(* Logix 5000 project; controller TFF vendor 1 type 14 code 107 rev 33.11; software revision 33.04; part 7 of 38 *)

        [4,11].DelayTimer.PRE := 2000, [4,11].DelayTimerSP := 2, [4,11].EnableCfg := 1, [4,11].ActiveStateCFg := 1, [4,11].RealInputCfg := 1, [4,11].InputAddressCfg := 11, [4,12].Tag := 'ZS007', [4,12].DelayTimer.PRE := 2000, [4,12].DelayTimerSP := 2, [4,12].EnableCfg := 1, [4,12].ActiveStateCFg := 1, [4,12].RealInputCfg := 1, [4,12].InputAddressCfg := 12, [4,13].Tag := 'ZS008', [4,13].AlarmCurrentValue := 1, [4,13].Override := 1, [4,13].DelayTimer.PRE := 20000, [4,13].DelayTimerSP := 2, [4,13].Priority := 1, [4,13].EnableCfg := 1, [4,13].ActiveStateCFg := 1, [4,13].RealInputCfg := 1, [4,13].InputAddressCfg := 13, [4,13].AlarmCfg := 1, [4,13].OverrideCfg := 1, [4,13].PriorityCfg := 1, [4,13].Cond1Cfg := 1, [4,14].Tag := 'XS011', [4,14].DelayTimer.PRE := 2000, [4,14].DelayTimerSP := 2, [4,14].EnableCfg := 1, [4,14].ActiveStateCFg := 1, [4,14].RealInputCfg := 1, [4,14].InputAddressCfg := 14, [4,15].Tag := 'XS012', [4,15].SoftInput := 1, [4,15].DelayTimer.PRE := 2000, [4,15].DelayTimerSP := 2, [4,15].EnableCfg := 1, [4,15].ActiveStateCFg := 1, [4,15].RealInputCfg := 1, [4,15].InputAddressCfg := 15, [4,16].Tag := 'SIC001DF', [4,16].AlarmCurrentValue := 1, [4,16].Override := 1, [4,16].SoftInput := 1, [4,16].DelayTimer.PRE := 1000, [4,16].DelayTimer.ACC := 3148, [4,16].DelayTimer.EN := 1, [4,16].DelayTimer.DN := 1, [4,16].DelayTimerSP := 1, [4,16].Priority := 1, [4,16].EnableCfg := 1, [4,16].ActiveStateCFg := 1, [4,16].RealInputCfg := 1, [4,16].InputAddressCfg := 16, [4,16].AlarmCfg := 1, [4,16].OverrideCfg := 1, [4,16].PriorityCfg := 1, [4,17].Tag := 'SIC002DF',
        [4,17].AlarmCurrentValue := 1, [4,17].Override := 1, [4,17].SoftInput := 1, [4,17].DelayTimer.PRE := 1000, [4,17].DelayTimer.ACC := 2449345, [4,17].DelayTimer.EN := 1, [4,17].DelayTimer.DN := 1, [4,17].DelayTimerSP := 1, [4,17].Priority := 1, [4,17].EnableCfg := 1, [4,17].ActiveStateCFg := 1, [4,17].RealInputCfg := 1, [4,17].InputAddressCfg := 17, [4,17].AlarmCfg := 1, [4,17].OverrideCfg := 1, [4,17].PriorityCfg := 1, [4,18].Tag := 'AA008', [4,18].AlarmCurrentValue := 1, [4,18].Override := 1, [4,18].DelayTimer.PRE := 1000, [4,18].DelayTimer.ACC := 1042, [4,18].DelayTimer.EN := 1, [4,18].DelayTimer.DN := 1, [4,18].DelayTimerSP := 1, [4,18].Priority := 1, [4,18].EnableCfg := 1, [4,18].ActiveStateCFg := 1, [4,18].RealInputCfg := 1, [4,18].InputAddressCfg := 18, [4,18].AlarmCfg := 1, [4,18].OverrideCfg := 1, [4,18].PriorityCfg := 1, [4,19].Tag := 'LSH001', [4,19].AlarmCurrentValue := 1, [4,19].Override := 1, [4,19].DelayTimer.PRE := 1000, [4,19].DelayTimer.EN := 1, [4,19].DelayTimer.DN := 1, [4,19].DelayTimerSP := 1, [4,19].EnableCfg := 1, [4,19].ActiveStateCFg := 1, [4,19].RealInputCfg := 1, [4,19].InputAddressCfg := 19, [4,19].AlarmCfg := 1, [4,19].OverrideCfg := 1, [4,19].PriorityCfg := 1, [4,20].Tag := 'LSL002', [4,20].AlarmCurrentValue := 1, [4,20].Override := 1, [4,20].DelayTimer.PRE := 1000, [4,20].DelayTimer.EN := 1, [4,20].DelayTimer.DN := 1, [4,20].DelayTimerSP := 1, [4,20].EnableCfg := 1, [4,20].ActiveStateCFg := 1, [4,20].RealInputCfg := 1, [4,20].InputAddressCfg := 20, [4,20].AlarmCfg := 1, [4,20].OverrideCfg := 1, [4,20].PriorityCfg := 1,
        [4,21].Tag := 'PSH001', [4,21].AlarmCurrentValue := 1, [4,21].AlarmAck := 1, [4,21].Alarm := 1, [4,21].Mimic := 5, [4,21].DelayTimer.PRE := 1000, [4,21].DelayTimer.ACC := 1042, [4,21].DelayTimer.EN := 1, [4,21].DelayTimer.DN := 1, [4,21].DelayTimerSP := 1, [4,21].Priority := 1, [4,21].EnableCfg := 1, [4,21].ActiveStateCFg := 1, [4,21].RealInputCfg := 1, [4,21].InputAddressCfg := 21, [4,21].AlarmCfg := 1, [4,21].AlarmONS := 1, [4,22].Tag := 'PSH002', [4,22].AlarmCurrentValue := 1, [4,22].AlarmAck := 1, [4,22].Alarm := 1, [4,22].Mimic := 5, [4,22].DelayTimer.PRE := 1000, [4,22].DelayTimer.ACC := 1042, [4,22].DelayTimer.EN := 1, [4,22].DelayTimer.DN := 1, [4,22].DelayTimerSP := 1, [4,22].Priority := 1, [4,22].EnableCfg := 1, [4,22].ActiveStateCFg := 1, [4,22].RealInputCfg := 1, [4,22].InputAddressCfg := 22, [4,22].AlarmCfg := 1, [4,22].AlarmONS := 1, [4,23].Tag := 'DF48VP001', [4,23].AlarmCurrentValue := 1, [4,23].Override := 1, [4,23].DelayTimer.PRE := 1000, [4,23].DelayTimer.ACC := 1042, [4,23].DelayTimer.EN := 1, [4,23].DelayTimer.DN := 1, [4,23].DelayTimerSP := 1, [4,23].Priority := 1, [4,23].EnableCfg := 1, [4,23].ActiveStateCFg := 1, [4,23].RealInputCfg := 1, [4,23].InputAddressCfg := 23, [4,23].AlarmCfg := 1, [4,23].OverrideCfg := 1, [4,23].PriorityCfg := 1, [4,24].Tag := 'DF48VP002', [4,24].AlarmCurrentValue := 1, [4,24].Override := 1, [4,24].DelayTimer.PRE := 1000, [4,24].DelayTimer.ACC := 1043, [4,24].DelayTimer.EN := 1, [4,24].DelayTimer.DN := 1, [4,24].DelayTimerSP := 1, [4,24].Priority := 1, [4,24].EnableCfg := 1,
        [4,24].ActiveStateCFg := 1, [4,24].RealInputCfg := 1, [4,24].InputAddressCfg := 24, [4,24].AlarmCfg := 1, [4,24].OverrideCfg := 1, [4,24].PriorityCfg := 1, [4,25].Tag := 'XS002', [4,25].AlarmCurrentValue := 1, [4,25].Override := 1, [4,25].DelayTimer.PRE := 20000, [4,25].DelayTimerSP := 2, [4,25].Priority := 1, [4,25].EnableCfg := 1, [4,25].ActiveStateCFg := 1, [4,25].RealInputCfg := 1, [4,25].InputAddressCfg := 25, [4,25].AlarmCfg := 1, [4,25].OverrideCfg := 1, [4,25].PriorityCfg := 1, [4,25].Cond1Cfg := 1, [4,26].Override := 1, [4,26].ActiveStateCFg := 1, [4,26].RealInputCfg := 1, [4,26].InputAddressCfg := 26, [4,26].OverrideCfg := 1, [4,26].PriorityCfg := 1, [4,27].Override := 1, [4,27].SoftInput := 1, [4,27].ActiveStateCFg := 1, [4,27].RealInputCfg := 1, [4,27].InputAddressCfg := 27, [4,27].OverrideCfg := 1, [4,27].PriorityCfg := 1, [4,28].Override := 1, [4,28].SoftInput := 1, [4,28].ActiveStateCFg := 1, [4,28].RealInputCfg := 1, [4,28].InputAddressCfg := 28, [4,28].OverrideCfg := 1, [4,28].PriorityCfg := 1, [4,29].Override := 1, [4,29].SoftInput := 1, [4,29].ActiveStateCFg := 1, [4,29].RealInputCfg := 1, [4,29].InputAddressCfg := 29, [4,29].OverrideCfg := 1, [4,29].PriorityCfg := 1, [4,30].Override := 1, [4,30].SoftInput := 1, [4,30].ActiveStateCFg := 1, [4,30].RealInputCfg := 1, [4,30].InputAddressCfg := 30, [4,30].OverrideCfg := 1, [4,30].PriorityCfg := 1, [4,31].Override := 1, [4,31].ActiveStateCFg := 1, [4,31].RealInputCfg := 1, [4,31].InputAddressCfg := 31, [4,31].OverrideCfg := 1, [4,31].PriorityCfg := 1,
        [4,34].Tag := 'DI1', [4,34].Override := 1, [4,34].SoftInput := 1, [4,34].EnableCfg := 1, [4,34].ActiveStateCFg := 1, [4,34].RealInputCfg := 1, [4,34].InputAddressCfg := 34, [4,34].OverrideCfg := 1, [4,34].PriorityCfg := 1, [4,35].Tag := 'DI2', [4,35].Override := 1, [4,35].EnableCfg := 1, [4,35].ActiveStateCFg := 1, [4,35].RealInputCfg := 1, [4,35].InputAddressCfg := 35, [4,35].OverrideCfg := 1, [4,35].PriorityCfg := 1, [4,36].Tag := 'DI3', [4,36].Override := 1, [4,36].SoftInput := 1, [4,36].EnableCfg := 1, [4,36].ActiveStateCFg := 1, [4,36].RealInputCfg := 1, [4,36].InputAddressCfg := 36, [4,36].OverrideCfg := 1, [4,36].PriorityCfg := 1, [4,37].Tag := 'DI4', [4,37].Override := 1, [4,37].EnableCfg := 1, [4,37].ActiveStateCFg := 1, [4,37].RealInputCfg := 1, [4,37].InputAddressCfg := 37, [4,37].OverrideCfg := 1, [4,37].PriorityCfg := 1, [4,38].Tag := 'DI5', [4,38].Override := 1, [4,38].EnableCfg := 1, [4,38].ActiveStateCFg := 1, [4,38].RealInputCfg := 1, [4,38].InputAddressCfg := 38, [4,38].OverrideCfg := 1, [4,38].PriorityCfg := 1, [4,39].Tag := 'DI6', [4,39].Override := 1, [4,39].SoftInput := 1, [4,39].EnableCfg := 1, [4,39].ActiveStateCFg := 1, [4,39].RealInputCfg := 1, [4,39].InputAddressCfg := 39, [4,39].OverrideCfg := 1, [4,39].PriorityCfg := 1, [4,40].Tag := 'DI7', [4,40].Override := 1, [4,40].EnableCfg := 1, [4,40].ActiveStateCFg := 1, [4,40].RealInputCfg := 1, [4,40].InputAddressCfg := 40, [4,40].OverrideCfg := 1, [4,40].PriorityCfg := 1, [4,41].Tag := 'DI8',
        [4,41].Override := 1, [4,41].EnableCfg := 1, [4,41].ActiveStateCFg := 1, [4,41].RealInputCfg := 1, [4,41].InputAddressCfg := 41, [4,41].OverrideCfg := 1, [4,41].PriorityCfg := 1, [4,50].Tag := 'YA01', [4,50].Desc := 'PC to PLC Com. Failure', [4,50].AlarmCurrentValue := 1, [4,50].Override := 1, [4,50].SoftInput := 1, [4,50].Condition1 := 1, [4,50].Cond1Text := 'HMI HeartBeat received', [4,50].DelayTimer.PRE := 60000, [4,50].DelayTimer.ACC := 598, [4,50].DelayTimer.EN := 1, [4,50].DelayTimer.TT := 1, [4,50].DelayTimerSP := 60, [4,50].EnableCfg := 1, [4,50].InputAddressCfg := 50, [4,50].AlarmCfg := 1, [4,50].AlarmStateCfg := 1, [4,50].OverrideCfg := 1, [4,50].PriorityCfg := 1, [4,50].Cond1Cfg := 1, [4,51].Tag := 'YA02', [4,51].Desc := 'CCP Runtime Com. Failure', [4,51].AlarmCurrentValue := 1, [4,51].Override := 1, [4,51].SoftInput := 1, [4,51].Condition1 := 1, [4,51].Cond1Text := 'HMI HeartBeat received', [4,51].DelayTimer.PRE := 60000, [4,51].DelayTimer.ACC := 60008, [4,51].DelayTimer.EN := 1, [4,51].DelayTimer.DN := 1, [4,51].DelayTimerSP := 60, [4,51].EnableCfg := 1, [4,51].InputAddressCfg := 51, [4,51].AlarmCfg := 1, [4,51].AlarmStateCfg := 1, [4,51].OverrideCfg := 1, [4,51].PriorityCfg := 1, [4,51].Cond1Cfg := 1, [4,52].Tag := 'YA03', [4,52].Desc := 'Hist. Data Collect. Fail', [4,52].AlarmCurrentValue := 1, [4,52].Override := 1, [4,52].SoftInput := 1, [4,52].Condition1 := 1, [4,52].Cond1Text := 'HMI HeartBeat received', [4,52].DelayTimer.PRE := 60000, [4,52].DelayTimer.ACC := 1145, [4,52].DelayTimer.EN := 1, [4,52].DelayTimer.TT := 1, [4,52].DelayTimerSP := 60, [4,52].EnableCfg := 1, [4,52].InputAddressCfg := 52, [4,52].AlarmCfg := 1,
        [4,52].AlarmStateCfg := 1, [4,52].OverrideCfg := 1, [4,52].PriorityCfg := 1, [4,52].Cond1Cfg := 1, [4,53].Tag := 'YA04', [4,53].Desc := 'HDD OverLoad', [4,53].Override := 1, [4,53].DelayTimer.PRE := 60000, [4,53].DelayTimerSP := 60, [4,53].EnableCfg := 1, [4,53].ActiveStateCFg := 1, [4,53].InputAddressCfg := 53, [4,53].AlarmCfg := 1, [4,53].AlarmStateCfg := 1, [4,53].OverrideCfg := 1, [4,53].PriorityCfg := 1, [4,54].Tag := 'YA05', [4,54].Override := 1, [4,54].DelayTimer.PRE := 60000, [4,54].DelayTimerSP := 60, [4,54].EnableCfg := 1, [4,54].ActiveStateCFg := 1, [4,54].InputAddressCfg := 54, [4,54].AlarmCfg := 1, [4,54].AlarmStateCfg := 1, [4,54].OverrideCfg := 1, [4,54].PriorityCfg := 1, [4,55].Tag := 'YA06', [4,55].CurrentValue := 1, [4,55].AlarmCurrentValue := 1, [4,55].Override := 1, [4,55].Mimic := 1, [4,55].SoftInput := 1, [4,55].DelayTimer.PRE := 5000, [4,55].DelayTimer.ACC := 5022, [4,55].DelayTimer.EN := 1, [4,55].DelayTimer.DN := 1, [4,55].DelayTimerSP := 5, [4,55].Priority := 1, [4,55].EnableCfg := 1, [4,55].ActiveStateCFg := 1, [4,55].InputAddressCfg := 55, [4,55].AlarmCfg := 1, [4,55].AlarmStateCfg := 1, [4,55].OverrideCfg := 1, [4,55].PriorityCfg := 1, [4,56].Tag := 'YA07', [4,56].CurrentValue := 1, [4,56].AlarmCurrentValue := 1, [4,56].Override := 1, [4,56].Mimic := 1, [4,56].SoftInput := 1, [4,56].DelayTimer.PRE := 2000, [4,56].DelayTimer.ACC := 2004, [4,56].DelayTimer.EN := 1, [4,56].DelayTimer.DN := 1, [4,56].DelayTimerSP := 2, [4,56].EnableCfg := 1, [4,56].ActiveStateCFg := 1, [4,56].InputAddressCfg := 56,
        [4,56].AlarmCfg := 1, [4,56].AlarmStateCfg := 1, [4,56].OverrideCfg := 1, [4,56].PriorityCfg := 1, [4,57].Tag := 'YA08', [4,57].CurrentValue := 1, [4,57].AlarmCurrentValue := 1, [4,57].Override := 1, [4,57].Mimic := 1, [4,57].SoftInput := 1, [4,57].DelayTimer.PRE := 5000, [4,57].DelayTimer.ACC := 5011, [4,57].DelayTimer.EN := 1, [4,57].DelayTimer.DN := 1, [4,57].DelayTimerSP := 5, [4,57].Priority := 1, [4,57].EnableCfg := 1, [4,57].ActiveStateCFg := 1, [4,57].InputAddressCfg := 57, [4,57].AlarmCfg := 1, [4,57].AlarmStateCfg := 1, [4,57].OverrideCfg := 1, [4,57].PriorityCfg := 1, [4,58].Tag := 'YA09', [4,58].CurrentValue := 1, [4,58].AlarmCurrentValue := 1, [4,58].Override := 1, [4,58].Mimic := 1, [4,58].SoftInput := 1, [4,58].DelayTimer.PRE := 2000, [4,58].DelayTimer.ACC := 2050, [4,58].DelayTimer.EN := 1, [4,58].DelayTimer.DN := 1, [4,58].DelayTimerSP := 2, [4,58].EnableCfg := 1, [4,58].ActiveStateCFg := 1, [4,58].InputAddressCfg := 58, [4,58].AlarmCfg := 1, [4,58].AlarmStateCfg := 1, [4,58].OverrideCfg := 1, [4,58].PriorityCfg := 1, [4,59].Tag := 'YA10', [4,59].CurrentValue := 1, [4,59].Mimic := 1, [4,59].Priority := 1, [4,59].EnableCfg := 1, [4,59].InputAddressCfg := 59, [4,59].AlarmCfg := 1, [4,59].AlarmStateCfg := 1, [4,60].Tag := 'YA11', [4,60].AlarmCurrentValue := 1, [4,60].Override := 1, [4,60].DelayTimer.PRE := 5000, [4,60].DelayTimer.ACC := 5010, [4,60].DelayTimer.EN := 1, [4,60].DelayTimer.DN := 1, [4,60].DelayTimerSP := 5, [4,60].EnableCfg := 1, [4,60].ActiveStateCFg := 1, [4,60].InputAddressCfg := 60,
        [4,60].AlarmCfg := 1, [4,60].OverrideCfg := 1, [4,60].PriorityCfg := 1, [4,61].Tag := 'YA12', [4,61].Override := 1, [4,61].DelayTimer.PRE := 2000, [4,61].DelayTimerSP := 2, [4,61].EnableCfg := 1, [4,61].ActiveStateCFg := 1, [4,61].InputAddressCfg := 61, [4,61].AlarmCfg := 1, [4,61].AlarmStateCfg := 1, [4,61].OverrideCfg := 1, [4,61].PriorityCfg := 1, [4,62].Tag := 'UserNCr1', [4,62].CurrentValue := 1, [4,62].Mimic := 1, [4,62].EnableCfg := 1, [4,62].InputAddressCfg := 62, [4,63].Tag := 'UserCr1', [4,63].SoftInput := 1, [4,63].Priority := 1, [4,63].EnableCfg := 1, [4,63].InputAddressCfg := 63, [4,64].Tag := 'UserNCr2', [4,64].CurrentValue := 1, [4,64].Mimic := 1, [4,64].EnableCfg := 1, [4,64].InputAddressCfg := 64, [4,65].Tag := 'UserCr2', [4,65].CurrentValue := 1, [4,65].Mimic := 1, [4,65].Priority := 1, [4,65].EnableCfg := 1, [4,65].InputAddressCfg := 65, [4,66].Tag := 'LV001_Err', [4,66].Override := 1, [4,66].DelayTimer.PRE := 2000, [4,66].DelayTimerSP := 2, [4,66].EnableCfg := 1, [4,66].ActiveStateCFg := 1, [4,66].InputAddressCfg := 66, [4,66].AlarmCfg := 1, [4,66].AlarmStateCfg := 1, [4,66].OverrideCfg := 1, [4,66].PriorityCfg := 1, [4,67].Tag := 'LV002_Err', [4,67].Override := 1, [4,67].DelayTimer.PRE := 2000, [4,67].DelayTimerSP := 2, [4,67].EnableCfg := 1, [4,67].ActiveStateCFg := 1, [4,67].InputAddressCfg := 67, [4,67].AlarmCfg := 1, [4,67].AlarmStateCfg := 1, [4,67].OverrideCfg := 1, [4,67].PriorityCfg := 1, [4,68].CurrentValue := 1, [4,68].AlarmCurrentValue := 1, [4,68].Override := 1,
        [4,68].Mimic := 1, [4,68].SoftInput := 1, [4,68].DelayTimer.PRE := 1000, [4,68].DelayTimer.ACC := 3526, [4,68].DelayTimer.EN := 1, [4,68].DelayTimer.DN := 1, [4,68].DelayTimerSP := 1, [4,68].Priority := 1, [4,68].EnableCfg := 1, [4,68].ActiveStateCFg := 1, [4,68].InputAddressCfg := 68, [4,68].AlarmCfg := 1, [4,68].AlarmStateCfg := 1, [4,68].OverrideCfg := 1, [4,69].Override := 1, [4,69].EnableCfg := 1, [4,69].ActiveStateCFg := 1, [4,69].InputAddressCfg := 69, [4,69].AlarmCfg := 1, [4,69].AlarmStateCfg := 1, [4,69].OverrideCfg := 1, [4,69].PriorityCfg := 1, [4,70].CurrentValue := 1, [4,70].Mimic := 1, [4,70].DelayTimer.PRE := 2000, [4,70].DelayTimerSP := 2, [4,70].Priority := 1, [4,70].ActiveStateCFg := 1, [4,70].InputAddressCfg := 70, [4,70].AlarmStateCfg := 1, [4,70].OverrideCfg := 1, [4,70].PriorityCfg := 1, [4,71].CurrentValue := 1, [4,71].AlarmCurrentValue := 1, [4,71].AlarmAck := 1, [4,71].Mimic := 5, [4,71].DelayTimer.PRE := 2000, [4,71].DelayTimer.ACC := 2053, [4,71].DelayTimer.EN := 1, [4,71].DelayTimer.DN := 1, [4,71].DelayTimerSP := 2, [4,71].Priority := 1, [4,71].ActiveStateCFg := 1, [4,71].InputAddressCfg := 71, [4,71].AlarmStateCfg := 1, [4,71].OverrideCfg := 1, [4,71].PriorityCfg := 1, [4,71].AlarmONS := 1, [4,72].CurrentValue := 1, [4,72].Mimic := 1, [4,72].DelayTimer.PRE := 2000, [4,72].DelayTimerSP := 2, [4,72].ActiveStateCFg := 1, [4,72].InputAddressCfg := 72, [4,72].AlarmStateCfg := 1, [4,72].OverrideCfg := 1, [4,72].PriorityCfg := 1, [4,73].CurrentValue := 1, [4,73].Mimic := 1, [4,73].DelayTimer.PRE := 2000,
        [4,73].DelayTimerSP := 2, [4,73].ActiveStateCFg := 1, [4,73].InputAddressCfg := 73, [4,73].AlarmStateCfg := 1, [4,73].OverrideCfg := 1, [4,73].PriorityCfg := 1, [4,74].CurrentValue := 1, [4,74].Mimic := 1, [4,74].DelayTimer.PRE := 2000, [4,74].DelayTimerSP := 2, [4,74].ActiveStateCFg := 1, [4,74].InputAddressCfg := 74, [4,74].AlarmStateCfg := 1, [4,74].OverrideCfg := 1, [4,74].PriorityCfg := 1, [4,75].CurrentValue := 1, [4,75].AlarmCurrentValue := 1, [4,75].AlarmAck := 1, [4,75].Alarm := 1, [4,75].Mimic := 3, [4,75].SoftInput := 1, [4,75].DelayTimer.PRE := 2000, [4,75].DelayTimer.ACC := 44, [4,75].DelayTimer.EN := 1, [4,75].DelayTimer.DN := 1, [4,75].DelayTimerSP := 2, [4,75].ActiveStateCFg := 1, [4,75].InputAddressCfg := 75, [4,75].AlarmStateCfg := 1, [4,75].OverrideCfg := 1, [4,75].PriorityCfg := 1, [4,75].AlarmONS := 1, [4,76].CurrentValue := 1, [4,76].Mimic := 1, [4,76].DelayTimer.PRE := 2000, [4,76].DelayTimerSP := 2, [4,76].Priority := 1, [4,76].ActiveStateCFg := 1, [4,76].InputAddressCfg := 76, [4,76].AlarmStateCfg := 1, [4,76].OverrideCfg := 1, [4,76].PriorityCfg := 1, [4,77].CurrentValue := 1, [4,77].Mimic := 1, [4,77].DelayTimer.PRE := 2000, [4,77].DelayTimerSP := 2, [4,77].Priority := 1, [4,77].ActiveStateCFg := 1, [4,77].InputAddressCfg := 77, [4,77].AlarmStateCfg := 1, [4,77].OverrideCfg := 1, [4,77].PriorityCfg := 1, [4,78].CurrentValue := 1, [4,78].AlarmCurrentValue := 1, [4,78].AlarmAck := 1, [4,78].Alarm := 1, [4,78].Mimic := 5, [4,78].SoftInput := 1, [4,78].DelayTimer.PRE := 2000, [4,78].DelayTimer.ACC := 45,
        [4,78].DelayTimer.EN := 1, [4,78].DelayTimer.DN := 1, [4,78].DelayTimerSP := 2, [4,78].Priority := 1, [4,78].ActiveStateCFg := 1, [4,78].InputAddressCfg := 78, [4,78].AlarmStateCfg := 1, [4,78].OverrideCfg := 1, [4,78].PriorityCfg := 1, [4,78].AlarmONS := 1, [4,79].CurrentValue := 1, [4,79].AlarmCurrentValue := 1, [4,79].Mimic := 1, [4,79].DelayTimer.PRE := 2000, [4,79].DelayTimer.ACC := 44, [4,79].DelayTimer.EN := 1, [4,79].DelayTimer.DN := 1, [4,79].DelayTimerSP := 2, [4,79].Priority := 1, [4,79].ActiveStateCFg := 1, [4,79].InputAddressCfg := 79, [4,79].AlarmStateCfg := 1, [4,79].OverrideCfg := 1, [4,79].PriorityCfg := 1, [4,80].CurrentValue := 1, [4,80].AlarmCurrentValue := 1, [4,80].Mimic := 1, [4,80].DelayTimer.PRE := 2000, [4,80].DelayTimer.ACC := 44, [4,80].DelayTimer.EN := 1, [4,80].DelayTimer.DN := 1, [4,80].DelayTimerSP := 2, [4,80].Priority := 1, [4,80].ActiveStateCFg := 1, [4,80].InputAddressCfg := 80, [4,80].AlarmStateCfg := 1, [4,80].OverrideCfg := 1, [4,80].PriorityCfg := 1, [4,81].CurrentValue := 1, [4,81].AlarmCurrentValue := 1, [4,81].Mimic := 1, [4,81].DelayTimer.PRE := 2000, [4,81].DelayTimer.ACC := 44, [4,81].DelayTimer.EN := 1, [4,81].DelayTimer.DN := 1, [4,81].DelayTimerSP := 2, [4,81].ActiveStateCFg := 1, [4,81].InputAddressCfg := 81, [4,81].AlarmStateCfg := 1, [4,81].OverrideCfg := 1, [4,81].PriorityCfg := 1, [4,82].CurrentValue := 1, [4,82].AlarmCurrentValue := 1, [4,82].Mimic := 1, [4,82].DelayTimer.PRE := 2000, [4,82].DelayTimer.ACC := 44, [4,82].DelayTimer.EN := 1, [4,82].DelayTimer.DN := 1, [4,82].DelayTimerSP := 2, [4,82].Priority := 1,
        [4,82].ActiveStateCFg := 1, [4,82].InputAddressCfg := 82, [4,82].AlarmStateCfg := 1, [4,82].OverrideCfg := 1, [4,82].PriorityCfg := 1, [4,83].CurrentValue := 1, [4,83].AlarmCurrentValue := 1, [4,83].AlarmAck := 1, [4,83].Alarm := 1, [4,83].Mimic := 5, [4,83].SoftInput := 1, [4,83].DelayTimer.PRE := 2000, [4,83].DelayTimer.ACC := 44, [4,83].DelayTimer.EN := 1, [4,83].DelayTimer.DN := 1, [4,83].DelayTimerSP := 2, [4,83].Priority := 1, [4,83].ActiveStateCFg := 1, [4,83].InputAddressCfg := 83, [4,83].AlarmStateCfg := 1, [4,83].OverrideCfg := 1, [4,83].PriorityCfg := 1, [4,83].AlarmONS := 1, [4,84].CurrentValue := 1, [4,84].Mimic := 1, [4,84].DelayTimer.PRE := 2000, [4,84].DelayTimerSP := 2, [4,84].Priority := 1, [4,84].ActiveStateCFg := 1, [4,84].InputAddressCfg := 84, [4,84].AlarmStateCfg := 1, [4,84].OverrideCfg := 1, [4,84].PriorityCfg := 1, [4,85].CurrentValue := 1, [4,85].AlarmCurrentValue := 1, [4,85].AlarmAck := 1, [4,85].Alarm := 1, [4,85].Mimic := 3, [4,85].SoftInput := 1, [4,85].DelayTimer.PRE := 2000, [4,85].DelayTimer.ACC := 2021, [4,85].DelayTimer.EN := 1, [4,85].DelayTimer.DN := 1, [4,85].DelayTimerSP := 2, [4,85].ActiveStateCFg := 1, [4,85].InputAddressCfg := 85, [4,85].AlarmStateCfg := 1, [4,85].OverrideCfg := 1, [4,85].PriorityCfg := 1, [4,85].AlarmONS := 1, [4,86].CurrentValue := 1, [4,86].Mimic := 1, [4,86].DelayTimer.PRE := 2000, [4,86].DelayTimerSP := 2, [4,86].ActiveStateCFg := 1, [4,86].InputAddressCfg := 86, [4,86].AlarmStateCfg := 1, [4,86].OverrideCfg := 1, [4,86].PriorityCfg := 1, [4,87].CurrentValue := 1,
        [4,87].Mimic := 1, [4,87].DelayTimer.PRE := 2000, [4,87].DelayTimerSP := 2, [4,87].ActiveStateCFg := 1, [4,87].InputAddressCfg := 87, [4,87].AlarmStateCfg := 1, [4,87].OverrideCfg := 1, [4,87].PriorityCfg := 1, [4,88].CurrentValue := 1, [4,88].Mimic := 1, [4,88].DelayTimer.PRE := 2000, [4,88].DelayTimerSP := 2, [4,88].ActiveStateCFg := 1, [4,88].InputAddressCfg := 88, [4,88].AlarmStateCfg := 1, [4,88].OverrideCfg := 1, [4,88].PriorityCfg := 1, [4,89].CurrentValue := 1, [4,89].Mimic := 1, [4,89].DelayTimer.PRE := 2000, [4,89].DelayTimerSP := 2, [4,89].ActiveStateCFg := 1, [4,89].InputAddressCfg := 89, [4,89].AlarmStateCfg := 1, [4,89].OverrideCfg := 1, [4,89].PriorityCfg := 1, [4,90].Tag := 'PI001_SIG', [4,90].CurrentValue := 1, [4,90].AlarmCurrentValue := 1, [4,90].AlarmAck := 1, [4,90].Alarm := 1, [4,90].Mimic := 5, [4,90].SoftInput := 1, [4,90].DelayTimer.PRE := 2000, [4,90].DelayTimer.ACC := 6308, [4,90].DelayTimer.EN := 1, [4,90].DelayTimer.DN := 1, [4,90].DelayTimerSP := 2, [4,90].Priority := 1, [4,90].EnableCfg := 1, [4,90].ActiveStateCFg := 1, [4,90].InputAddressCfg := 90, [4,90].AlarmCfg := 1, [4,90].AlarmStateCfg := 1, [4,90].OverrideCfg := 1, [4,90].PriorityCfg := 1, [4,90].AlarmONS := 1, [4,91].Tag := 'FI001_SIG', [4,91].CurrentValue := 1, [4,91].AlarmCurrentValue := 1, [4,91].AlarmAck := 1, [4,91].Alarm := 1, [4,91].Mimic := 5, [4,91].SoftInput := 1, [4,91].DelayTimer.PRE := 2000, [4,91].DelayTimer.ACC := 2025, [4,91].DelayTimer.EN := 1, [4,91].DelayTimer.DN := 1, [4,91].DelayTimerSP := 2, [4,91].Priority := 1,
        [4,91].EnableCfg := 1, [4,91].ActiveStateCFg := 1, [4,91].InputAddressCfg := 91, [4,91].AlarmCfg := 1, [4,91].AlarmStateCfg := 1, [4,91].OverrideCfg := 1, [4,91].PriorityCfg := 1, [4,91].AlarmONS := 1, [4,92].Tag := 'PI002_SIG', [4,92].CurrentValue := 1, [4,92].AlarmCurrentValue := 1, [4,92].AlarmAck := 1, [4,92].Alarm := 1, [4,92].Mimic := 5, [4,92].SoftInput := 1, [4,92].DelayTimer.PRE := 2000, [4,92].DelayTimer.EN := 1, [4,92].DelayTimer.DN := 1, [4,92].DelayTimerSP := 2, [4,92].Priority := 1, [4,92].EnableCfg := 1, [4,92].ActiveStateCFg := 1, [4,92].InputAddressCfg := 92, [4,92].AlarmCfg := 1, [4,92].AlarmStateCfg := 1, [4,92].OverrideCfg := 1, [4,92].PriorityCfg := 1, [4,92].AlarmONS := 1, [4,93].Tag := 'FI002_SIG', [4,93].CurrentValue := 1, [4,93].AlarmCurrentValue := 1, [4,93].AlarmAck := 1, [4,93].Alarm := 1, [4,93].Mimic := 5, [4,93].SoftInput := 1, [4,93].DelayTimer.PRE := 2000, [4,93].DelayTimer.ACC := 2049, [4,93].DelayTimer.EN := 1, [4,93].DelayTimer.DN := 1, [4,93].DelayTimerSP := 2, [4,93].Priority := 1, [4,93].EnableCfg := 1, [4,93].ActiveStateCFg := 1, [4,93].InputAddressCfg := 93, [4,93].AlarmCfg := 1, [4,93].AlarmStateCfg := 1, [4,93].OverrideCfg := 1, [4,93].PriorityCfg := 1, [4,93].AlarmONS := 1, [4,94].Tag := 'PI003_SIG', [4,94].CurrentValue := 1, [4,94].AlarmCurrentValue := 1, [4,94].AlarmAck := 1, [4,94].Alarm := 1, [4,94].Mimic := 3, [4,94].SoftInput := 1, [4,94].DelayTimer.PRE := 2000, [4,94].DelayTimer.ACC := 37, [4,94].DelayTimer.EN := 1, [4,94].DelayTimer.DN := 1,
        [4,94].DelayTimerSP := 2, [4,94].EnableCfg := 1, [4,94].ActiveStateCFg := 1, [4,94].InputAddressCfg := 94, [4,94].AlarmCfg := 1, [4,94].AlarmStateCfg := 1, [4,94].OverrideCfg := 1, [4,94].PriorityCfg := 1, [4,94].AlarmONS := 1, [4,95].Tag := 'AI102_SIG', [4,95].CurrentValue := 1, [4,95].AlarmCurrentValue := 1, [4,95].AlarmAck := 1, [4,95].Alarm := 1, [4,95].Mimic := 5, [4,95].SoftInput := 1, [4,95].DelayTimer.PRE := 2000, [4,95].DelayTimer.ACC := 3550, [4,95].DelayTimer.EN := 1, [4,95].DelayTimer.DN := 1, [4,95].DelayTimerSP := 2, [4,95].Priority := 1, [4,95].EnableCfg := 1, [4,95].ActiveStateCFg := 1, [4,95].InputAddressCfg := 95, [4,95].AlarmCfg := 1, [4,95].AlarmStateCfg := 1, [4,95].OverrideCfg := 1, [4,95].PriorityCfg := 1, [4,95].AlarmONS := 1, [4,96].Tag := 'AI103_SIG', [4,96].CurrentValue := 1, [4,96].AlarmCurrentValue := 1, [4,96].AlarmAck := 1, [4,96].Alarm := 1, [4,96].Mimic := 5, [4,96].SoftInput := 1, [4,96].DelayTimer.PRE := 2000, [4,96].DelayTimer.EN := 1, [4,96].DelayTimer.DN := 1, [4,96].DelayTimerSP := 2, [4,96].Priority := 1, [4,96].EnableCfg := 1, [4,96].ActiveStateCFg := 1, [4,96].InputAddressCfg := 96, [4,96].AlarmCfg := 1, [4,96].AlarmStateCfg := 1, [4,96].OverrideCfg := 1, [4,96].PriorityCfg := 1, [4,96].AlarmONS := 1, [4,97].Tag := 'AI201A_SIG', [4,97].CurrentValue := 1, [4,97].AlarmCurrentValue := 1, [4,97].AlarmAck := 1, [4,97].Alarm := 1, [4,97].Mimic := 5, [4,97].SoftInput := 1, [4,97].DelayTimer.PRE := 2000, [4,97].DelayTimer.EN := 1, [4,97].DelayTimer.DN := 1,
        [4,97].DelayTimerSP := 2, [4,97].Priority := 1, [4,97].EnableCfg := 1, [4,97].ActiveStateCFg := 1, [4,97].InputAddressCfg := 97, [4,97].AlarmCfg := 1, [4,97].AlarmStateCfg := 1, [4,97].OverrideCfg := 1, [4,97].PriorityCfg := 1, [4,97].AlarmONS := 1, [4,98].Tag := 'AI201B_SIG', [4,98].CurrentValue := 1, [4,98].AlarmCurrentValue := 1, [4,98].AlarmAck := 1, [4,98].Alarm := 1, [4,98].Mimic := 5, [4,98].SoftInput := 1, [4,98].DelayTimer.PRE := 2000, [4,98].DelayTimer.EN := 1, [4,98].DelayTimer.DN := 1, [4,98].DelayTimerSP := 2, [4,98].Priority := 1, [4,98].EnableCfg := 1, [4,98].ActiveStateCFg := 1, [4,98].InputAddressCfg := 98, [4,98].AlarmCfg := 1, [4,98].AlarmStateCfg := 1, [4,98].OverrideCfg := 1, [4,98].PriorityCfg := 1, [4,98].AlarmONS := 1, [4,99].Tag := 'TI201_SIG', [4,99].CurrentValue := 1, [4,99].AlarmCurrentValue := 1, [4,99].AlarmAck := 1, [4,99].Alarm := 1, [4,99].Mimic := 3, [4,99].SoftInput := 1, [4,99].DelayTimer.PRE := 2000, [4,99].DelayTimer.EN := 1, [4,99].DelayTimer.DN := 1, [4,99].DelayTimerSP := 2, [4,99].EnableCfg := 1, [4,99].ActiveStateCFg := 1, [4,99].InputAddressCfg := 99, [4,99].AlarmCfg := 1, [4,99].AlarmStateCfg := 1, [4,99].OverrideCfg := 1, [4,99].PriorityCfg := 1, [4,99].AlarmONS := 1, [4,100].Tag := 'AI202_SIG', [4,100].CurrentValue := 1, [4,100].AlarmCurrentValue := 1, [4,100].AlarmAck := 1, [4,100].Alarm := 1, [4,100].Mimic := 5, [4,100].SoftInput := 1, [4,100].DelayTimer.PRE := 2000, [4,100].DelayTimer.EN := 1, [4,100].DelayTimer.DN := 1, [4,100].DelayTimerSP := 2,
        [4,100].Priority := 1, [4,100].EnableCfg := 1, [4,100].ActiveStateCFg := 1, [4,100].InputAddressCfg := 100, [4,100].AlarmCfg := 1, [4,100].AlarmStateCfg := 1, [4,100].OverrideCfg := 1, [4,100].PriorityCfg := 1, [4,100].AlarmONS := 1, [4,101].Tag := 'AI203_SIG', [4,101].CurrentValue := 1, [4,101].AlarmCurrentValue := 1, [4,101].AlarmAck := 1, [4,101].Alarm := 1, [4,101].Mimic := 5, [4,101].SoftInput := 1, [4,101].DelayTimer.PRE := 2000, [4,101].DelayTimer.EN := 1, [4,101].DelayTimer.DN := 1, [4,101].DelayTimerSP := 2, [4,101].Priority := 1, [4,101].EnableCfg := 1, [4,101].ActiveStateCFg := 1, [4,101].InputAddressCfg := 101, [4,101].AlarmCfg := 1, [4,101].AlarmStateCfg := 1, [4,101].OverrideCfg := 1, [4,101].PriorityCfg := 1, [4,101].AlarmONS := 1, [4,102].Tag := 'AI204_SIG', [4,102].CurrentValue := 1, [4,102].AlarmCurrentValue := 1, [4,102].AlarmAck := 1, [4,102].Alarm := 1, [4,102].Mimic := 5, [4,102].SoftInput := 1, [4,102].DelayTimer.PRE := 2000, [4,102].DelayTimer.EN := 1, [4,102].DelayTimer.DN := 1, [4,102].DelayTimerSP := 2, [4,102].Priority := 1, [4,102].EnableCfg := 1, [4,102].ActiveStateCFg := 1, [4,102].InputAddressCfg := 102, [4,102].AlarmCfg := 1, [4,102].AlarmStateCfg := 1, [4,102].OverrideCfg := 1, [4,102].PriorityCfg := 1, [4,102].AlarmONS := 1, [4,103].Tag := 'PCV032_SIG', [4,103].CurrentValue := 1, [4,103].AlarmCurrentValue := 1, [4,103].AlarmAck := 1, [4,103].Alarm := 1, [4,103].Mimic := 5, [4,103].SoftInput := 1, [4,103].DelayTimer.PRE := 2000, [4,103].DelayTimer.ACC := 4119948, [4,103].DelayTimer.EN := 1, [4,103].DelayTimer.DN := 1,
        [4,103].DelayTimerSP := 2, [4,103].Priority := 1, [4,103].EnableCfg := 1, [4,103].ActiveStateCFg := 1, [4,103].InputAddressCfg := 103, [4,103].AlarmCfg := 1, [4,103].AlarmStateCfg := 1, [4,103].OverrideCfg := 1, [4,103].PriorityCfg := 1, [4,103].AlarmONS := 1, [5,0].Tag := 'PISL601', [5,0].AlarmCurrentValue := 1, [5,0].Override := 1, [5,0].DelayTimer.PRE := 2000, [5,0].DelayTimer.ACC := 129444, [5,0].DelayTimer.EN := 1, [5,0].DelayTimer.DN := 1, [5,0].DelayTimerSP := 2, [5,0].Priority := 1, [5,0].EnableCfg := 1, [5,0].ActiveStateCFg := 1, [5,0].RealInputCfg := 1, [5,0].AlarmCfg := 1, [5,0].OverrideCfg := 1, [5,0].PriorityCfg := 1, [5,1].Tag := 'PISL602', [5,1].AlarmCurrentValue := 1, [5,1].Override := 1, [5,1].Condition2 := 1, [5,1].DelayTimer.PRE := 2000, [5,1].DelayTimer.ACC := 44686, [5,1].DelayTimer.EN := 1, [5,1].DelayTimer.DN := 1, [5,1].DelayTimerSP := 2, [5,1].Priority := 1, [5,1].EnableCfg := 1, [5,1].ActiveStateCFg := 1, [5,1].RealInputCfg := 1, [5,1].InputAddressCfg := 1, [5,1].AlarmCfg := 1, [5,1].OverrideCfg := 1, [5,1].PriorityCfg := 1, [5,2].Tag := 'ES001', [5,2].CurrentValue := 1, [5,2].Mimic := 1, [5,2].DelayTimer.PRE := 1000, [5,2].DelayTimerSP := 1, [5,2].Priority := 1, [5,2].EnableCfg := 1, [5,2].ActiveStateCFg := 1, [5,2].RealInputCfg := 1, [5,2].InputAddressCfg := 2, [5,2].AlarmCfg := 1, [5,3].Tag := 'RSBUZZ', [5,3].DelayTimer.PRE := 2000, [5,3].DelayTimerSP := 2, [5,3].EnableCfg := 1, [5,3].ActiveStateCFg := 1, [5,3].RealInputCfg := 1, [5,3].InputAddressCfg := 3,
        [5,4].Tag := 'DF24VDC', [5,4].AlarmCurrentValue := 1, [5,4].Override := 1, [5,4].DelayTimer.PRE := 1000, [5,4].DelayTimer.ACC := 11063, [5,4].DelayTimer.EN := 1, [5,4].DelayTimer.DN := 1, [5,4].DelayTimerSP := 1, [5,4].Priority := 1, [5,4].EnableCfg := 1, [5,4].ActiveStateCFg := 1, [5,4].RealInputCfg := 1, [5,4].InputAddressCfg := 4, [5,4].AlarmCfg := 1, [5,4].OverrideCfg := 1, [5,4].PriorityCfg := 1, [5,5].Tag := 'ZS008', [5,5].AlarmCurrentValue := 1, [5,5].Override := 1, [5,5].DelayTimer.PRE := 1000, [5,5].DelayTimer.ACC := 1072, [5,5].DelayTimer.EN := 1, [5,5].DelayTimer.DN := 1, [5,5].DelayTimerSP := 1, [5,5].Priority := 1, [5,5].EnableCfg := 1, [5,5].ActiveStateCFg := 1, [5,5].RealInputCfg := 1, [5,5].InputAddressCfg := 5, [5,5].AlarmCfg := 1, [5,5].OverrideCfg := 1, [5,6].Tag := 'ZS001', [5,6].DelayTimer.PRE := 2000, [5,6].DelayTimerSP := 2, [5,6].EnableCfg := 1, [5,6].ActiveStateCFg := 1, [5,6].RealInputCfg := 1, [5,6].InputAddressCfg := 6, [5,7].Tag := 'ZS002', [5,7].DelayTimer.PRE := 2000, [5,7].DelayTimerSP := 2, [5,7].EnableCfg := 1, [5,7].ActiveStateCFg := 1, [5,7].RealInputCfg := 1, [5,7].InputAddressCfg := 7, [5,8].Tag := 'ZS003', [5,8].DelayTimer.PRE := 2000, [5,8].DelayTimerSP := 2, [5,8].EnableCfg := 1, [5,8].ActiveStateCFg := 1, [5,8].RealInputCfg := 1, [5,8].InputAddressCfg := 8, [5,9].Tag := 'ZS004', [5,9].DelayTimer.PRE := 2000, [5,9].DelayTimerSP := 2, [5,9].EnableCfg := 1, [5,9].ActiveStateCFg := 1, [5,9].RealInputCfg := 1, [5,9].InputAddressCfg := 9, [5,10].Tag := 'ZS005',
        [5,10].DelayTimer.PRE := 2000, [5,10].DelayTimerSP := 2, [5,10].EnableCfg := 1, [5,10].ActiveStateCFg := 1, [5,10].RealInputCfg := 1, [5,10].InputAddressCfg := 10, [5,11].Tag := 'ZS006', [5,11].DelayTimer.PRE := 2000, [5,11].DelayTimerSP := 2, [5,11].EnableCfg := 1, [5,11].ActiveStateCFg := 1, [5,11].RealInputCfg := 1, [5,11].InputAddressCfg := 11, [5,12].Tag := 'ZS007', [5,12].DelayTimer.PRE := 2000, [5,12].DelayTimerSP := 2, [5,12].EnableCfg := 1, [5,12].ActiveStateCFg := 1, [5,12].RealInputCfg := 1, [5,12].InputAddressCfg := 12, [5,13].Tag := 'ZS008', [5,13].AlarmCurrentValue := 1, [5,13].Override := 1, [5,13].DelayTimer.PRE := 20000, [5,13].DelayTimerSP := 2, [5,13].Priority := 1, [5,13].EnableCfg := 1, [5,13].ActiveStateCFg := 1, [5,13].RealInputCfg := 1, [5,13].InputAddressCfg := 13, [5,13].AlarmCfg := 1, [5,13].OverrideCfg := 1, [5,13].PriorityCfg := 1, [5,13].Cond1Cfg := 1, [5,14].Tag := 'XS011', [5,14].DelayTimer.PRE := 2000, [5,14].DelayTimerSP := 2, [5,14].EnableCfg := 1, [5,14].ActiveStateCFg := 1, [5,14].RealInputCfg := 1, [5,14].InputAddressCfg := 14, [5,15].Tag := 'XS012', [5,15].SoftInput := 1, [5,15].DelayTimer.PRE := 2000, [5,15].DelayTimerSP := 2, [5,15].EnableCfg := 1, [5,15].ActiveStateCFg := 1, [5,15].RealInputCfg := 1, [5,15].InputAddressCfg := 15, [5,16].Tag := 'SIC001DF', [5,16].AlarmCurrentValue := 1, [5,16].Override := 1, [5,16].SoftInput := 1, [5,16].DelayTimer.PRE := 1000, [5,16].DelayTimer.ACC := 3148, [5,16].DelayTimer.EN := 1, [5,16].DelayTimer.DN := 1, [5,16].DelayTimerSP := 1, [5,16].Priority := 1, [5,16].EnableCfg := 1,
        [5,16].ActiveStateCFg := 1, [5,16].RealInputCfg := 1, [5,16].InputAddressCfg := 16, [5,16].AlarmCfg := 1, [5,16].OverrideCfg := 1, [5,16].PriorityCfg := 1, [5,17].Tag := 'SIC002DF', [5,17].AlarmCurrentValue := 1, [5,17].Override := 1, [5,17].SoftInput := 1, [5,17].DelayTimer.PRE := 1000, [5,17].DelayTimer.ACC := 2449345, [5,17].DelayTimer.EN := 1, [5,17].DelayTimer.DN := 1, [5,17].DelayTimerSP := 1, [5,17].Priority := 1, [5,17].EnableCfg := 1, [5,17].ActiveStateCFg := 1, [5,17].RealInputCfg := 1, [5,17].InputAddressCfg := 17, [5,17].AlarmCfg := 1, [5,17].OverrideCfg := 1, [5,17].PriorityCfg := 1, [5,18].Tag := 'AA008', [5,18].AlarmCurrentValue := 1, [5,18].Override := 1, [5,18].DelayTimer.PRE := 1000, [5,18].DelayTimer.EN := 1, [5,18].DelayTimer.DN := 1, [5,18].DelayTimerSP := 1, [5,18].Priority := 1, [5,18].EnableCfg := 1, [5,18].ActiveStateCFg := 1, [5,18].RealInputCfg := 1, [5,18].InputAddressCfg := 18, [5,18].AlarmCfg := 1, [5,18].OverrideCfg := 1, [5,18].PriorityCfg := 1, [5,19].Tag := 'LSH001', [5,19].AlarmCurrentValue := 1, [5,19].Override := 1, [5,19].DelayTimer.PRE := 1000, [5,19].DelayTimer.EN := 1, [5,19].DelayTimer.DN := 1, [5,19].DelayTimerSP := 1, [5,19].EnableCfg := 1, [5,19].ActiveStateCFg := 1, [5,19].RealInputCfg := 1, [5,19].InputAddressCfg := 19, [5,19].AlarmCfg := 1, [5,19].OverrideCfg := 1, [5,19].PriorityCfg := 1, [5,20].Tag := 'LSL002', [5,20].AlarmCurrentValue := 1, [5,20].Override := 1, [5,20].DelayTimer.PRE := 1000, [5,20].DelayTimer.EN := 1, [5,20].DelayTimer.DN := 1, [5,20].DelayTimerSP := 1, [5,20].EnableCfg := 1,
        [5,20].ActiveStateCFg := 1, [5,20].RealInputCfg := 1, [5,20].InputAddressCfg := 20, [5,20].AlarmCfg := 1, [5,20].OverrideCfg := 1, [5,20].PriorityCfg := 1, [5,21].Tag := 'PSH001', [5,21].AlarmCurrentValue := 1, [5,21].AlarmAck := 1, [5,21].Alarm := 1, [5,21].Mimic := 5, [5,21].DelayTimer.PRE := 1000, [5,21].DelayTimer.ACC := 44686, [5,21].DelayTimer.EN := 1, [5,21].DelayTimer.DN := 1, [5,21].DelayTimerSP := 1, [5,21].Priority := 1, [5,21].EnableCfg := 1, [5,21].ActiveStateCFg := 1, [5,21].RealInputCfg := 1, [5,21].InputAddressCfg := 21, [5,21].AlarmCfg := 1, [5,21].AlarmONS := 1, [5,22].Tag := 'PSH002', [5,22].AlarmCurrentValue := 1, [5,22].AlarmAck := 1, [5,22].Alarm := 1, [5,22].Mimic := 5, [5,22].DelayTimer.PRE := 1000, [5,22].DelayTimer.ACC := 44686, [5,22].DelayTimer.EN := 1, [5,22].DelayTimer.DN := 1, [5,22].DelayTimerSP := 1, [5,22].Priority := 1, [5,22].EnableCfg := 1, [5,22].ActiveStateCFg := 1, [5,22].RealInputCfg := 1, [5,22].InputAddressCfg := 22, [5,22].AlarmCfg := 1, [5,22].AlarmONS := 1, [5,23].Tag := 'DF48VP001', [5,23].AlarmCurrentValue := 1, [5,23].Override := 1, [5,23].DelayTimer.PRE := 1000, [5,23].DelayTimer.ACC := 3043, [5,23].DelayTimer.EN := 1, [5,23].DelayTimer.DN := 1, [5,23].DelayTimerSP := 1, [5,23].Priority := 1, [5,23].EnableCfg := 1, [5,23].ActiveStateCFg := 1, [5,23].RealInputCfg := 1, [5,23].InputAddressCfg := 23, [5,23].AlarmCfg := 1, [5,23].OverrideCfg := 1, [5,23].PriorityCfg := 1, [5,24].Tag := 'DF48VP002', [5,24].AlarmCurrentValue := 1, [5,24].Override := 1, [5,24].DelayTimer.PRE := 1000,
        [5,24].DelayTimer.EN := 1, [5,24].DelayTimer.DN := 1, [5,24].DelayTimerSP := 1, [5,24].Priority := 1, [5,24].EnableCfg := 1, [5,24].ActiveStateCFg := 1, [5,24].RealInputCfg := 1, [5,24].InputAddressCfg := 24, [5,24].AlarmCfg := 1, [5,24].OverrideCfg := 1, [5,24].PriorityCfg := 1, [5,25].Tag := 'XS002', [5,25].AlarmCurrentValue := 1, [5,25].Override := 1, [5,25].DelayTimer.PRE := 20000, [5,25].DelayTimerSP := 2, [5,25].Priority := 1, [5,25].EnableCfg := 1, [5,25].ActiveStateCFg := 1, [5,25].RealInputCfg := 1, [5,25].InputAddressCfg := 25, [5,25].AlarmCfg := 1, [5,25].OverrideCfg := 1, [5,25].PriorityCfg := 1, [5,25].Cond1Cfg := 1, [5,26].Override := 1, [5,26].ActiveStateCFg := 1, [5,26].RealInputCfg := 1, [5,26].InputAddressCfg := 26, [5,26].OverrideCfg := 1, [5,26].PriorityCfg := 1, [5,27].Override := 1, [5,27].SoftInput := 1, [5,27].ActiveStateCFg := 1, [5,27].RealInputCfg := 1, [5,27].InputAddressCfg := 27, [5,27].OverrideCfg := 1, [5,27].PriorityCfg := 1, [5,28].Override := 1, [5,28].SoftInput := 1, [5,28].ActiveStateCFg := 1, [5,28].RealInputCfg := 1, [5,28].InputAddressCfg := 28, [5,28].OverrideCfg := 1, [5,28].PriorityCfg := 1, [5,29].Override := 1, [5,29].SoftInput := 1, [5,29].ActiveStateCFg := 1, [5,29].RealInputCfg := 1, [5,29].InputAddressCfg := 29, [5,29].OverrideCfg := 1, [5,29].PriorityCfg := 1, [5,30].Override := 1, [5,30].SoftInput := 1, [5,30].ActiveStateCFg := 1, [5,30].RealInputCfg := 1, [5,30].InputAddressCfg := 30, [5,30].OverrideCfg := 1, [5,30].PriorityCfg := 1, [5,31].Override := 1,
        [5,31].ActiveStateCFg := 1, [5,31].RealInputCfg := 1, [5,31].InputAddressCfg := 31, [5,31].OverrideCfg := 1, [5,31].PriorityCfg := 1, [5,34].Tag := 'DI1', [5,34].Override := 1, [5,34].SoftInput := 1, [5,34].EnableCfg := 1, [5,34].ActiveStateCFg := 1, [5,34].RealInputCfg := 1, [5,34].InputAddressCfg := 34, [5,34].OverrideCfg := 1, [5,34].PriorityCfg := 1, [5,35].Tag := 'DI2', [5,35].Override := 1, [5,35].EnableCfg := 1, [5,35].ActiveStateCFg := 1, [5,35].RealInputCfg := 1, [5,35].InputAddressCfg := 35, [5,35].OverrideCfg := 1, [5,35].PriorityCfg := 1, [5,36].Tag := 'DI3', [5,36].Override := 1, [5,36].SoftInput := 1, [5,36].EnableCfg := 1, [5,36].ActiveStateCFg := 1, [5,36].RealInputCfg := 1, [5,36].InputAddressCfg := 36, [5,36].OverrideCfg := 1, [5,36].PriorityCfg := 1, [5,37].Tag := 'DI4', [5,37].Override := 1, [5,37].EnableCfg := 1, [5,37].ActiveStateCFg := 1, [5,37].RealInputCfg := 1, [5,37].InputAddressCfg := 37, [5,37].OverrideCfg := 1, [5,37].PriorityCfg := 1, [5,38].Tag := 'DI5', [5,38].Override := 1, [5,38].EnableCfg := 1, [5,38].ActiveStateCFg := 1, [5,38].RealInputCfg := 1, [5,38].InputAddressCfg := 38, [5,38].OverrideCfg := 1, [5,38].PriorityCfg := 1, [5,39].Tag := 'DI6', [5,39].Override := 1, [5,39].SoftInput := 1, [5,39].EnableCfg := 1, [5,39].ActiveStateCFg := 1, [5,39].RealInputCfg := 1, [5,39].InputAddressCfg := 39, [5,39].OverrideCfg := 1, [5,39].PriorityCfg := 1, [5,40].Tag := 'DI7', [5,40].Override := 1, [5,40].EnableCfg := 1, [5,40].ActiveStateCFg := 1,
        [5,40].RealInputCfg := 1, [5,40].InputAddressCfg := 40, [5,40].OverrideCfg := 1, [5,40].PriorityCfg := 1, [5,41].Tag := 'DI8', [5,41].Override := 1, [5,41].EnableCfg := 1, [5,41].ActiveStateCFg := 1, [5,41].RealInputCfg := 1, [5,41].InputAddressCfg := 41, [5,41].OverrideCfg := 1, [5,41].PriorityCfg := 1, [5,50].Tag := 'YA01', [5,50].Desc := 'PC to PLC Com. Failure', [5,50].AlarmCurrentValue := 1, [5,50].Override := 1, [5,50].SoftInput := 1, [5,50].Cond1Text := 'HMI HeartBeat received', [5,50].DelayTimer.PRE := 60000, [5,50].DelayTimerSP := 60, [5,50].EnableCfg := 1, [5,50].InputAddressCfg := 50, [5,50].AlarmCfg := 1, [5,50].AlarmStateCfg := 1, [5,50].OverrideCfg := 1, [5,50].PriorityCfg := 1, [5,50].Cond1Cfg := 1, [5,51].Tag := 'YA02', [5,51].Desc := 'CCP Runtime Com. Failure', [5,51].AlarmCurrentValue := 1, [5,51].Override := 1, [5,51].SoftInput := 1, [5,51].Cond1Text := 'HMI HeartBeat received', [5,51].DelayTimer.PRE := 60000, [5,51].DelayTimerSP := 60, [5,51].EnableCfg := 1, [5,51].InputAddressCfg := 51, [5,51].AlarmCfg := 1, [5,51].AlarmStateCfg := 1, [5,51].OverrideCfg := 1, [5,51].PriorityCfg := 1, [5,51].Cond1Cfg := 1, [5,52].Tag := 'YA03', [5,52].Desc := 'Hist. Data Collect. Fail', [5,52].AlarmCurrentValue := 1, [5,52].Override := 1, [5,52].SoftInput := 1, [5,52].Cond1Text := 'HMI HeartBeat received', [5,52].DelayTimer.PRE := 60000, [5,52].DelayTimerSP := 60, [5,52].EnableCfg := 1, [5,52].InputAddressCfg := 52, [5,52].AlarmCfg := 1, [5,52].AlarmStateCfg := 1, [5,52].OverrideCfg := 1, [5,52].PriorityCfg := 1, [5,52].Cond1Cfg := 1, [5,53].Tag := 'YA04', [5,53].Desc := 'HDD OverLoad', [5,53].Override := 1,
        [5,53].DelayTimer.PRE := 60000, [5,53].DelayTimerSP := 60, [5,53].EnableCfg := 1, [5,53].ActiveStateCFg := 1, [5,53].InputAddressCfg := 53, [5,53].AlarmCfg := 1, [5,53].AlarmStateCfg := 1, [5,53].OverrideCfg := 1, [5,53].PriorityCfg := 1, [5,54].Tag := 'YA05', [5,54].Override := 1, [5,54].DelayTimer.PRE := 60000, [5,54].DelayTimerSP := 60, [5,54].EnableCfg := 1, [5,54].ActiveStateCFg := 1, [5,54].InputAddressCfg := 54, [5,54].AlarmCfg := 1, [5,54].AlarmStateCfg := 1, [5,54].OverrideCfg := 1, [5,54].PriorityCfg := 1, [5,55].Tag := 'YA06', [5,55].CurrentValue := 1, [5,55].AlarmCurrentValue := 1, [5,55].Override := 1, [5,55].Mimic := 1, [5,55].SoftInput := 1, [5,55].DelayTimer.PRE := 5000, [5,55].DelayTimer.ACC := 36135, [5,55].DelayTimer.EN := 1, [5,55].DelayTimer.DN := 1, [5,55].DelayTimerSP := 5, [5,55].Priority := 1, [5,55].EnableCfg := 1, [5,55].ActiveStateCFg := 1, [5,55].InputAddressCfg := 55, [5,55].AlarmCfg := 1, [5,55].AlarmStateCfg := 1, [5,55].OverrideCfg := 1, [5,55].PriorityCfg := 1, [5,56].Tag := 'YA07', [5,56].Override := 1, [5,56].DelayTimer.PRE := 2000, [5,56].DelayTimerSP := 2, [5,56].EnableCfg := 1, [5,56].ActiveStateCFg := 1, [5,56].InputAddressCfg := 56, [5,56].AlarmCfg := 1, [5,56].AlarmStateCfg := 1, [5,56].OverrideCfg := 1, [5,56].PriorityCfg := 1, [5,57].Tag := 'YA08', [5,57].CurrentValue := 1, [5,57].AlarmCurrentValue := 1, [5,57].Override := 1, [5,57].Mimic := 1, [5,57].SoftInput := 1, [5,57].DelayTimer.PRE := 5000, [5,57].DelayTimer.ACC := 1036, [5,57].DelayTimer.EN := 1, [5,57].DelayTimer.DN := 1,
        [5,57].DelayTimerSP := 5, [5,57].Priority := 1, [5,57].EnableCfg := 1, [5,57].ActiveStateCFg := 1, [5,57].InputAddressCfg := 57, [5,57].AlarmCfg := 1, [5,57].AlarmStateCfg := 1, [5,57].OverrideCfg := 1, [5,57].PriorityCfg := 1, [5,58].Tag := 'YA09', [5,58].Override := 1, [5,58].DelayTimer.PRE := 2000, [5,58].DelayTimerSP := 2, [5,58].EnableCfg := 1, [5,58].ActiveStateCFg := 1, [5,58].InputAddressCfg := 58, [5,58].AlarmCfg := 1, [5,58].AlarmStateCfg := 1, [5,58].OverrideCfg := 1, [5,58].PriorityCfg := 1, [5,59].Tag := 'YA10', [5,59].CurrentValue := 1, [5,59].Mimic := 1, [5,59].Priority := 1, [5,59].EnableCfg := 1, [5,59].InputAddressCfg := 59, [5,59].AlarmCfg := 1, [5,59].AlarmStateCfg := 1, [5,60].Tag := 'YA11', [5,60].AlarmCurrentValue := 1, [5,60].Override := 1, [5,60].DelayTimer.PRE := 5000, [5,60].DelayTimer.ACC := 2469476, [5,60].DelayTimer.EN := 1, [5,60].DelayTimer.DN := 1, [5,60].DelayTimerSP := 5, [5,60].EnableCfg := 1, [5,60].ActiveStateCFg := 1, [5,60].InputAddressCfg := 60, [5,60].AlarmCfg := 1, [5,60].OverrideCfg := 1, [5,60].PriorityCfg := 1, [5,61].Tag := 'YA12', [5,61].Override := 1, [5,61].DelayTimer.PRE := 2000, [5,61].DelayTimerSP := 2, [5,61].EnableCfg := 1, [5,61].ActiveStateCFg := 1, [5,61].InputAddressCfg := 61, [5,61].AlarmCfg := 1, [5,61].AlarmStateCfg := 1, [5,61].OverrideCfg := 1, [5,61].PriorityCfg := 1, [5,62].Tag := 'UserNCr1', [5,62].CurrentValue := 1, [5,62].Mimic := 1, [5,62].EnableCfg := 1, [5,62].InputAddressCfg := 62, [5,63].Tag := 'UserCr1', [5,63].CurrentValue := 1,
        [5,63].Mimic := 1, [5,63].Priority := 1, [5,63].EnableCfg := 1, [5,63].InputAddressCfg := 63, [5,64].Tag := 'UserNCr2', [5,64].CurrentValue := 1, [5,64].Mimic := 1, [5,64].EnableCfg := 1, [5,64].InputAddressCfg := 64, [5,65].Tag := 'UserCr2', [5,65].CurrentValue := 1, [5,65].Mimic := 1, [5,65].Priority := 1, [5,65].EnableCfg := 1, [5,65].InputAddressCfg := 65, [5,66].Tag := 'LV001_Err', [5,66].Override := 1, [5,66].DelayTimer.PRE := 2000, [5,66].DelayTimerSP := 2, [5,66].EnableCfg := 1, [5,66].ActiveStateCFg := 1, [5,66].InputAddressCfg := 66, [5,66].AlarmCfg := 1, [5,66].AlarmStateCfg := 1, [5,66].OverrideCfg := 1, [5,66].PriorityCfg := 1, [5,67].Tag := 'LV002_Err', [5,67].Override := 1, [5,67].DelayTimer.PRE := 2000, [5,67].DelayTimerSP := 2, [5,67].EnableCfg := 1, [5,67].ActiveStateCFg := 1, [5,67].InputAddressCfg := 67, [5,67].AlarmCfg := 1, [5,67].AlarmStateCfg := 1, [5,67].OverrideCfg := 1, [5,67].PriorityCfg := 1, [5,68].CurrentValue := 1, [5,68].AlarmCurrentValue := 1, [5,68].Override := 1, [5,68].Mimic := 1, [5,68].SoftInput := 1, [5,68].DelayTimer.PRE := 1000, [5,68].DelayTimer.ACC := 3526, [5,68].DelayTimer.EN := 1, [5,68].DelayTimer.DN := 1, [5,68].DelayTimerSP := 1, [5,68].Priority := 1, [5,68].EnableCfg := 1, [5,68].ActiveStateCFg := 1, [5,68].InputAddressCfg := 68, [5,68].AlarmCfg := 1, [5,68].AlarmStateCfg := 1, [5,68].OverrideCfg := 1, [5,69].CurrentValue := 1, [5,69].AlarmCurrentValue := 1, [5,69].AlarmAck := 1, [5,69].Alarm := 1, [5,69].Mimic := 5, [5,69].SoftInput := 1,
        [5,69].DelayTimer.PRE := 2000, [5,69].DelayTimer.ACC := 2052, [5,69].DelayTimer.EN := 1, [5,69].DelayTimer.DN := 1, [5,69].DelayTimerSP := 2, [5,69].Priority := 1, [5,69].ActiveStateCFg := 1, [5,69].InputAddressCfg := 69, [5,69].AlarmStateCfg := 1, [5,69].OverrideCfg := 1, [5,69].PriorityCfg := 1, [5,69].AlarmONS := 1, [5,70].CurrentValue := 1, [5,70].Mimic := 1, [5,70].DelayTimer.PRE := 2000, [5,70].DelayTimerSP := 2, [5,70].Priority := 1, [5,70].ActiveStateCFg := 1, [5,70].InputAddressCfg := 70, [5,70].AlarmStateCfg := 1, [5,70].OverrideCfg := 1, [5,70].PriorityCfg := 1, [5,71].CurrentValue := 1, [5,71].AlarmCurrentValue := 1, [5,71].AlarmAck := 1, [5,71].Mimic := 5, [5,71].DelayTimer.PRE := 2000, [5,71].DelayTimer.ACC := 2053, [5,71].DelayTimer.EN := 1, [5,71].DelayTimer.DN := 1, [5,71].DelayTimerSP := 2, [5,71].Priority := 1, [5,71].ActiveStateCFg := 1, [5,71].InputAddressCfg := 71, [5,71].AlarmStateCfg := 1, [5,71].OverrideCfg := 1, [5,71].PriorityCfg := 1, [5,71].AlarmONS := 1, [5,72].CurrentValue := 1, [5,72].Mimic := 1, [5,72].DelayTimer.PRE := 2000, [5,72].DelayTimerSP := 2, [5,72].ActiveStateCFg := 1, [5,72].InputAddressCfg := 72, [5,72].AlarmStateCfg := 1, [5,72].OverrideCfg := 1, [5,72].PriorityCfg := 1, [5,73].CurrentValue := 1, [5,73].Mimic := 1, [5,73].DelayTimer.PRE := 2000, [5,73].DelayTimerSP := 2, [5,73].ActiveStateCFg := 1, [5,73].InputAddressCfg := 73, [5,73].AlarmStateCfg := 1, [5,73].OverrideCfg := 1, [5,73].PriorityCfg := 1, [5,74].CurrentValue := 1, [5,74].Mimic := 1, [5,74].DelayTimer.PRE := 2000, [5,74].DelayTimerSP := 2,
        [5,74].ActiveStateCFg := 1, [5,74].InputAddressCfg := 74, [5,74].AlarmStateCfg := 1, [5,74].OverrideCfg := 1, [5,74].PriorityCfg := 1, [5,75].CurrentValue := 1, [5,75].AlarmCurrentValue := 1, [5,75].AlarmAck := 1, [5,75].Alarm := 1, [5,75].Mimic := 3, [5,75].SoftInput := 1, [5,75].DelayTimer.PRE := 2000, [5,75].DelayTimer.ACC := 44, [5,75].DelayTimer.EN := 1, [5,75].DelayTimer.DN := 1, [5,75].DelayTimerSP := 2, [5,75].ActiveStateCFg := 1, [5,75].InputAddressCfg := 75, [5,75].AlarmStateCfg := 1, [5,75].OverrideCfg := 1, [5,75].PriorityCfg := 1, [5,75].AlarmONS := 1, [5,76].CurrentValue := 1, [5,76].Mimic := 1, [5,76].DelayTimer.PRE := 2000, [5,76].DelayTimerSP := 2, [5,76].Priority := 1, [5,76].ActiveStateCFg := 1, [5,76].InputAddressCfg := 76, [5,76].AlarmStateCfg := 1, [5,76].OverrideCfg := 1, [5,76].PriorityCfg := 1, [5,77].CurrentValue := 1, [5,77].Mimic := 1, [5,77].DelayTimer.PRE := 2000, [5,77].DelayTimerSP := 2, [5,77].Priority := 1, [5,77].ActiveStateCFg := 1, [5,77].InputAddressCfg := 77, [5,77].AlarmStateCfg := 1, [5,77].OverrideCfg := 1, [5,77].PriorityCfg := 1, [5,78].CurrentValue := 1, [5,78].AlarmCurrentValue := 1, [5,78].AlarmAck := 1, [5,78].Alarm := 1, [5,78].Mimic := 5, [5,78].SoftInput := 1, [5,78].DelayTimer.PRE := 2000, [5,78].DelayTimer.ACC := 45, [5,78].DelayTimer.EN := 1, [5,78].DelayTimer.DN := 1, [5,78].DelayTimerSP := 2, [5,78].Priority := 1, [5,78].ActiveStateCFg := 1, [5,78].InputAddressCfg := 78, [5,78].AlarmStateCfg := 1, [5,78].OverrideCfg := 1, [5,78].PriorityCfg := 1, [5,78].AlarmONS := 1,
        [5,79].CurrentValue := 1, [5,79].AlarmCurrentValue := 1, [5,79].Mimic := 1, [5,79].DelayTimer.PRE := 2000, [5,79].DelayTimer.ACC := 44, [5,79].DelayTimer.EN := 1, [5,79].DelayTimer.DN := 1, [5,79].DelayTimerSP := 2, [5,79].Priority := 1, [5,79].ActiveStateCFg := 1, [5,79].InputAddressCfg := 79, [5,79].AlarmStateCfg := 1, [5,79].OverrideCfg := 1, [5,79].PriorityCfg := 1, [5,80].CurrentValue := 1, [5,80].AlarmCurrentValue := 1, [5,80].Mimic := 1, [5,80].DelayTimer.PRE := 2000, [5,80].DelayTimer.ACC := 44, [5,80].DelayTimer.EN := 1, [5,80].DelayTimer.DN := 1, [5,80].DelayTimerSP := 2, [5,80].Priority := 1, [5,80].ActiveStateCFg := 1, [5,80].InputAddressCfg := 80, [5,80].AlarmStateCfg := 1, [5,80].OverrideCfg := 1, [5,80].PriorityCfg := 1, [5,81].CurrentValue := 1, [5,81].AlarmCurrentValue := 1, [5,81].Mimic := 1, [5,81].DelayTimer.PRE := 2000, [5,81].DelayTimer.ACC := 44, [5,81].DelayTimer.EN := 1, [5,81].DelayTimer.DN := 1, [5,81].DelayTimerSP := 2, [5,81].ActiveStateCFg := 1, [5,81].InputAddressCfg := 81, [5,81].AlarmStateCfg := 1, [5,81].OverrideCfg := 1, [5,81].PriorityCfg := 1, [5,82].CurrentValue := 1, [5,82].AlarmCurrentValue := 1, [5,82].Mimic := 1, [5,82].DelayTimer.PRE := 2000, [5,82].DelayTimer.ACC := 44, [5,82].DelayTimer.EN := 1, [5,82].DelayTimer.DN := 1, [5,82].DelayTimerSP := 2, [5,82].Priority := 1, [5,82].ActiveStateCFg := 1, [5,82].InputAddressCfg := 82, [5,82].AlarmStateCfg := 1, [5,82].OverrideCfg := 1, [5,82].PriorityCfg := 1, [5,83].CurrentValue := 1, [5,83].AlarmCurrentValue := 1, [5,83].AlarmAck := 1, [5,83].Alarm := 1, [5,83].Mimic := 5,
        [5,83].SoftInput := 1, [5,83].DelayTimer.PRE := 2000, [5,83].DelayTimer.ACC := 44, [5,83].DelayTimer.EN := 1, [5,83].DelayTimer.DN := 1, [5,83].DelayTimerSP := 2, [5,83].Priority := 1, [5,83].ActiveStateCFg := 1, [5,83].InputAddressCfg := 83, [5,83].AlarmStateCfg := 1, [5,83].OverrideCfg := 1, [5,83].PriorityCfg := 1, [5,83].AlarmONS := 1, [5,84].CurrentValue := 1, [5,84].Mimic := 1, [5,84].DelayTimer.PRE := 2000, [5,84].DelayTimerSP := 2, [5,84].Priority := 1, [5,84].ActiveStateCFg := 1, [5,84].InputAddressCfg := 84, [5,84].AlarmStateCfg := 1, [5,84].OverrideCfg := 1, [5,84].PriorityCfg := 1, [5,85].CurrentValue := 1, [5,85].AlarmCurrentValue := 1, [5,85].AlarmAck := 1, [5,85].Alarm := 1, [5,85].Mimic := 3, [5,85].SoftInput := 1, [5,85].DelayTimer.PRE := 2000, [5,85].DelayTimer.ACC := 2021, [5,85].DelayTimer.EN := 1, [5,85].DelayTimer.DN := 1, [5,85].DelayTimerSP := 2, [5,85].ActiveStateCFg := 1, [5,85].InputAddressCfg := 85, [5,85].AlarmStateCfg := 1, [5,85].OverrideCfg := 1, [5,85].PriorityCfg := 1, [5,85].AlarmONS := 1, [5,86].CurrentValue := 1, [5,86].Mimic := 1, [5,86].DelayTimer.PRE := 2000, [5,86].DelayTimerSP := 2, [5,86].ActiveStateCFg := 1, [5,86].InputAddressCfg := 86, [5,86].AlarmStateCfg := 1, [5,86].OverrideCfg := 1, [5,86].PriorityCfg := 1, [5,87].CurrentValue := 1, [5,87].Mimic := 1, [5,87].DelayTimer.PRE := 2000, [5,87].DelayTimerSP := 2, [5,87].ActiveStateCFg := 1, [5,87].InputAddressCfg := 87, [5,87].AlarmStateCfg := 1, [5,87].OverrideCfg := 1, [5,87].PriorityCfg := 1, [5,88].CurrentValue := 1, [5,88].Mimic := 1,
        [5,88].DelayTimer.PRE := 2000, [5,88].DelayTimerSP := 2, [5,88].ActiveStateCFg := 1, [5,88].InputAddressCfg := 88, [5,88].AlarmStateCfg := 1, [5,88].OverrideCfg := 1, [5,88].PriorityCfg := 1, [5,89].CurrentValue := 1, [5,89].Mimic := 1, [5,89].DelayTimer.PRE := 2000, [5,89].DelayTimerSP := 2, [5,89].ActiveStateCFg := 1, [5,89].InputAddressCfg := 89, [5,89].AlarmStateCfg := 1, [5,89].OverrideCfg := 1, [5,89].PriorityCfg := 1, [5,90].Tag := 'PI001_SIG', [5,90].CurrentValue := 1, [5,90].AlarmCurrentValue := 1, [5,90].Override := 1, [5,90].Mimic := 1, [5,90].SoftInput := 1, [5,90].DelayTimer.PRE := 2000, [5,90].DelayTimer.ACC := 6308, [5,90].DelayTimer.EN := 1, [5,90].DelayTimer.DN := 1, [5,90].DelayTimerSP := 2, [5,90].Priority := 1, [5,90].EnableCfg := 1, [5,90].ActiveStateCFg := 1, [5,90].InputAddressCfg := 90, [5,90].AlarmCfg := 1, [5,90].AlarmStateCfg := 1, [5,90].OverrideCfg := 1, [5,90].PriorityCfg := 1, [5,91].Tag := 'FI001_SIG', [5,91].Override := 1, [5,91].DelayTimer.PRE := 2000, [5,91].DelayTimerSP := 2, [5,91].Priority := 1, [5,91].EnableCfg := 1, [5,91].ActiveStateCFg := 1, [5,91].InputAddressCfg := 91, [5,91].AlarmCfg := 1, [5,91].AlarmStateCfg := 1, [5,91].OverrideCfg := 1, [5,91].PriorityCfg := 1, [5,92].Tag := 'PI002_SIG', [5,92].CurrentValue := 1, [5,92].AlarmCurrentValue := 1, [5,92].Override := 1, [5,92].Mimic := 1, [5,92].SoftInput := 1, [5,92].DelayTimer.PRE := 2000, [5,92].DelayTimer.EN := 1, [5,92].DelayTimer.DN := 1, [5,92].DelayTimerSP := 2, [5,92].Priority := 1, [5,92].EnableCfg := 1, [5,92].ActiveStateCFg := 1,
        [5,92].InputAddressCfg := 92, [5,92].AlarmCfg := 1, [5,92].AlarmStateCfg := 1, [5,92].OverrideCfg := 1, [5,92].PriorityCfg := 1, [5,93].Tag := 'FI002_SIG', [5,93].Override := 1, [5,93].DelayTimer.PRE := 2000, [5,93].DelayTimerSP := 2, [5,93].Priority := 1, [5,93].EnableCfg := 1, [5,93].ActiveStateCFg := 1, [5,93].InputAddressCfg := 93, [5,93].AlarmCfg := 1, [5,93].AlarmStateCfg := 1, [5,93].OverrideCfg := 1, [5,93].PriorityCfg := 1, [5,94].Tag := 'PI003_SIG', [5,94].CurrentValue := 1, [5,94].AlarmCurrentValue := 1, [5,94].Override := 1, [5,94].Mimic := 1, [5,94].SoftInput := 1, [5,94].DelayTimer.PRE := 2000, [5,94].DelayTimer.ACC := 37, [5,94].DelayTimer.EN := 1, [5,94].DelayTimer.DN := 1, [5,94].DelayTimerSP := 2, [5,94].EnableCfg := 1, [5,94].ActiveStateCFg := 1, [5,94].InputAddressCfg := 94, [5,94].AlarmCfg := 1, [5,94].AlarmStateCfg := 1, [5,94].OverrideCfg := 1, [5,94].PriorityCfg := 1, [5,95].Tag := 'AI102_SIG', [5,95].CurrentValue := 1, [5,95].AlarmCurrentValue := 1, [5,95].Override := 1, [5,95].Mimic := 1, [5,95].SoftInput := 1, [5,95].DelayTimer.PRE := 2000, [5,95].DelayTimer.ACC := 3550, [5,95].DelayTimer.EN := 1, [5,95].DelayTimer.DN := 1, [5,95].DelayTimerSP := 2, [5,95].Priority := 1, [5,95].EnableCfg := 1, [5,95].ActiveStateCFg := 1, [5,95].InputAddressCfg := 95, [5,95].AlarmCfg := 1, [5,95].AlarmStateCfg := 1, [5,95].OverrideCfg := 1, [5,95].PriorityCfg := 1, [5,96].Tag := 'AI103_SIG', [5,96].CurrentValue := 1, [5,96].AlarmCurrentValue := 1, [5,96].Override := 1, [5,96].Mimic := 1, [5,96].SoftInput := 1,
        [5,96].DelayTimer.PRE := 2000, [5,96].DelayTimer.EN := 1, [5,96].DelayTimer.DN := 1, [5,96].DelayTimerSP := 2, [5,96].Priority := 1, [5,96].EnableCfg := 1, [5,96].ActiveStateCFg := 1, [5,96].InputAddressCfg := 96, [5,96].AlarmCfg := 1, [5,96].AlarmStateCfg := 1, [5,96].OverrideCfg := 1, [5,96].PriorityCfg := 1, [5,97].Tag := 'AI201A_SIG', [5,97].CurrentValue := 1, [5,97].AlarmCurrentValue := 1, [5,97].Override := 1, [5,97].Mimic := 1, [5,97].SoftInput := 1, [5,97].DelayTimer.PRE := 2000, [5,97].DelayTimer.EN := 1, [5,97].DelayTimer.DN := 1, [5,97].DelayTimerSP := 2, [5,97].Priority := 1, [5,97].EnableCfg := 1, [5,97].ActiveStateCFg := 1, [5,97].InputAddressCfg := 97, [5,97].AlarmCfg := 1, [5,97].AlarmStateCfg := 1, [5,97].OverrideCfg := 1, [5,97].PriorityCfg := 1, [5,98].Tag := 'AI201B_SIG', [5,98].CurrentValue := 1, [5,98].AlarmCurrentValue := 1, [5,98].Override := 1, [5,98].Mimic := 1, [5,98].SoftInput := 1, [5,98].DelayTimer.PRE := 2000, [5,98].DelayTimer.EN := 1, [5,98].DelayTimer.DN := 1, [5,98].DelayTimerSP := 2, [5,98].Priority := 1, [5,98].EnableCfg := 1, [5,98].ActiveStateCFg := 1, [5,98].InputAddressCfg := 98, [5,98].AlarmCfg := 1, [5,98].AlarmStateCfg := 1, [5,98].OverrideCfg := 1, [5,98].PriorityCfg := 1, [5,99].Tag := 'TI201_SIG', [5,99].CurrentValue := 1, [5,99].AlarmCurrentValue := 1, [5,99].Override := 1, [5,99].Mimic := 1, [5,99].SoftInput := 1, [5,99].DelayTimer.PRE := 2000, [5,99].DelayTimer.EN := 1, [5,99].DelayTimer.DN := 1, [5,99].DelayTimerSP := 2, [5,99].EnableCfg := 1, [5,99].ActiveStateCFg := 1,
        [5,99].InputAddressCfg := 99, [5,99].AlarmCfg := 1, [5,99].AlarmStateCfg := 1, [5,99].OverrideCfg := 1, [5,99].PriorityCfg := 1, [5,100].Tag := 'AI202_SIG', [5,100].CurrentValue := 1, [5,100].AlarmCurrentValue := 1, [5,100].Override := 1, [5,100].Mimic := 1, [5,100].SoftInput := 1, [5,100].DelayTimer.PRE := 2000, [5,100].DelayTimer.EN := 1, [5,100].DelayTimer.DN := 1, [5,100].DelayTimerSP := 2, [5,100].Priority := 1, [5,100].EnableCfg := 1, [5,100].ActiveStateCFg := 1, [5,100].InputAddressCfg := 100, [5,100].AlarmCfg := 1, [5,100].AlarmStateCfg := 1, [5,100].OverrideCfg := 1, [5,100].PriorityCfg := 1, [5,101].Tag := 'AI203_SIG', [5,101].CurrentValue := 1, [5,101].AlarmCurrentValue := 1, [5,101].Override := 1, [5,101].Mimic := 1, [5,101].SoftInput := 1, [5,101].DelayTimer.PRE := 2000, [5,101].DelayTimer.EN := 1, [5,101].DelayTimer.DN := 1, [5,101].DelayTimerSP := 2, [5,101].Priority := 1, [5,101].EnableCfg := 1, [5,101].ActiveStateCFg := 1, [5,101].InputAddressCfg := 101, [5,101].AlarmCfg := 1, [5,101].AlarmStateCfg := 1, [5,101].OverrideCfg := 1, [5,101].PriorityCfg := 1, [5,102].Tag := 'AI204_SIG', [5,102].CurrentValue := 1, [5,102].AlarmCurrentValue := 1, [5,102].Override := 1, [5,102].Mimic := 1, [5,102].SoftInput := 1, [5,102].DelayTimer.PRE := 2000, [5,102].DelayTimer.EN := 1, [5,102].DelayTimer.DN := 1, [5,102].DelayTimerSP := 2, [5,102].Priority := 1, [5,102].EnableCfg := 1, [5,102].ActiveStateCFg := 1, [5,102].InputAddressCfg := 102, [5,102].AlarmCfg := 1, [5,102].AlarmStateCfg := 1, [5,102].OverrideCfg := 1, [5,102].PriorityCfg := 1, [5,103].Tag := 'PCV032_SIG',
        [5,103].CurrentValue := 1, [5,103].AlarmCurrentValue := 1, [5,103].Override := 1, [5,103].Mimic := 1, [5,103].SoftInput := 1, [5,103].DelayTimer.PRE := 2000, [5,103].DelayTimer.EN := 1, [5,103].DelayTimer.DN := 1, [5,103].DelayTimerSP := 2, [5,103].Priority := 1, [5,103].EnableCfg := 1, [5,103].ActiveStateCFg := 1, [5,103].InputAddressCfg := 103, [5,103].AlarmCfg := 1, [5,103].AlarmStateCfg := 1, [5,103].OverrideCfg := 1, [5,103].PriorityCfg := 1);
   DO1 : ALIAS FOR DigitalOutput[80];
   DO2 : ALIAS FOR DigitalOutput[81];
   DO3 : ALIAS FOR DigitalOutput[82];
   DO4 : ALIAS FOR DigitalOutput[83];
   DO5 : ALIAS FOR DigitalOutput[84];
   DO6 : ALIAS FOR DigitalOutput[85];
   DO7 : ALIAS FOR DigitalOutput[86];
   DP : ALIAS FOR AnalogPoint[40];
   DPAlarm : ALIAS FOR AlarmAnalog[40];
   Drive : Drive[11] := ([0].InterlockTimer.ACC := 583, [0].InterlockTimer.EN := 1, [0].InterlockTimer.DN := 1, [1].TagName := 'SIC001', [1].RunInterlock := 1, [1].OutputAddress := 15, [1].InterlockTimer.PRE := 1000, [1].InterlockTimer.ACC := 1054, [1].InterlockTimer.EN := 1, [1].InterlockTimer.DN := 1, [1].EnableCfg := 1, [1].DriveStatus := 1, [2].TagName := 'SIC002', [2].RunInterlock := 1, [2].OutputAddress := 9, [2].InterlockTimer.PRE := 1000, [2].InterlockTimer.ACC := 1054, [2].InterlockTimer.EN := 1, [2].InterlockTimer.DN := 1, [2].EnableCfg := 1, [2].DriveStatus := 1, [3].TagName := 'SIC003', [3].RunInterlock := 1, [3].OutputAddress := 16, [3].InterlockTimer.PRE := 1000, [3].InterlockTimer.ACC := 1054, [3].InterlockTimer.EN := 1, [3].InterlockTimer.DN := 1, [3].EnableCfg := 1, [3].DriveStatus := 1, [5].RunOns := 1, [5].StopOns := 1);   // Drives Array
        [1]   // Feed Pump
        [2]   // Transfer Pump
        [3]   // Mixer
   Drive_Storage : Drive[6,11] := ([0,0].InterlockTimer.ACC := 583, [0,0].InterlockTimer.EN := 1, [0,0].InterlockTimer.DN := 1, [0,1].TagName := 'P001', [0,1].Desc := 'Primary Feed Pump', [0,1].RunInterlock := 1, [0,1].OutputAddress := 8, [0,1].InterlockTimer.PRE := 1000, [0,1].InterlockTimer.ACC := 1066, [0,1].InterlockTimer.EN := 1, [0,1].InterlockTimer.DN := 1, [0,1].EnableCfg := 1, [0,1].DriveStatus := 1, [0,1].DriveAlarmStatus := 2, [0,2].TagName := 'P002', [0,2].Desc := 'Secondary Feed Pump', [0,2].RunInterlock := 1, [0,2].OutputAddress := 9, [0,2].InterlockTimer.PRE := 1000, [0,2].InterlockTimer.ACC := 1066, [0,2].InterlockTimer.EN := 1, [0,2].InterlockTimer.DN := 1, [0,2].EnableCfg := 1, [0,2].DriveStatus := 1, [0,2].DriveAlarmStatus := 2, [0,5].RunOns := 1, [0,5].StopOns := 1, [1,0].InterlockTimer.ACC := 583, [1,0].InterlockTimer.EN := 1, [1,0].InterlockTimer.DN := 1, [1,1].TagName := 'P001', [1,1].Desc := 'Primary Feed Pump', [1,1].RunInterlock := 1, [1,1].OutputAddress := 8, [1,1].InterlockTimer.PRE := 1000, [1,1].InterlockTimer.ACC := 1066, [1,1].InterlockTimer.EN := 1, [1,1].InterlockTimer.DN := 1, [1,1].EnableCfg := 1, [1,1].DriveStatus := 1, [1,1].DriveAlarmStatus := 2, [1,2].TagName := 'P002', [1,2].Desc := 'Secondary Feed Pump', [1,2].RunInterlock := 1, [1,2].OutputAddress := 9, [1,2].InterlockTimer.PRE := 1000, [1,2].InterlockTimer.ACC := 1066, [1,2].InterlockTimer.EN := 1, [1,2].InterlockTimer.DN := 1, [1,2].EnableCfg := 1, [1,2].DriveStatus := 1, [1,2].DriveAlarmStatus := 2, [1,5].RunOns := 1, [1,5].StopOns := 1, [2,0].InterlockTimer.ACC := 583, [2,0].InterlockTimer.EN := 1, [2,0].InterlockTimer.DN := 1, [2,1].TagName := 'P001', [2,1].Desc := 'Primary Feed Pump', [2,1].RunInterlock := 1,
        [2,1].OutputAddress := 8, [2,1].InterlockTimer.PRE := 1000, [2,1].InterlockTimer.ACC := 1066, [2,1].InterlockTimer.EN := 1, [2,1].InterlockTimer.DN := 1, [2,1].EnableCfg := 1, [2,1].DriveStatus := 1, [2,1].DriveAlarmStatus := 2, [2,2].TagName := 'P002', [2,2].Desc := 'Secondary Feed Pump', [2,2].RunInterlock := 1, [2,2].OutputAddress := 9, [2,2].InterlockTimer.PRE := 1000, [2,2].InterlockTimer.ACC := 1066, [2,2].InterlockTimer.EN := 1, [2,2].InterlockTimer.DN := 1, [2,2].EnableCfg := 1, [2,2].DriveStatus := 1, [2,2].DriveAlarmStatus := 2, [2,5].RunOns := 1, [2,5].StopOns := 1, [3,1].RunInterlock := 1, [3,1].OutputAddress := 8, [3,1].InterlockTimer.PRE := 1000, [3,1].InterlockTimer.ACC := 134082, [3,1].InterlockTimer.EN := 1, [3,1].InterlockTimer.DN := 1, [3,1].EnableCfg := 1, [3,1].DriveStatus := 1, [3,1].DriveAlarmStatus := 1, [3,2].RunInterlock := 1, [3,2].OutputAddress := 9, [3,2].InterlockTimer.PRE := 1000, [3,2].InterlockTimer.ACC := 134082, [3,2].InterlockTimer.EN := 1, [3,2].InterlockTimer.DN := 1, [3,2].EnableCfg := 1, [3,2].DriveStatus := 1, [3,2].DriveAlarmStatus := 1, [4,0].InterlockTimer.ACC := 583, [4,0].InterlockTimer.EN := 1, [4,0].InterlockTimer.DN := 1, [4,1].TagName := 'P001', [4,1].Desc := 'Primary Feed Pump', [4,1].RunInterlock := 1, [4,1].OutputAddress := 8, [4,1].InterlockTimer.PRE := 1000, [4,1].InterlockTimer.ACC := 1097, [4,1].InterlockTimer.EN := 1, [4,1].InterlockTimer.DN := 1, [4,1].EnableCfg := 1, [4,1].DriveStatus := 1, [4,2].TagName := 'P002', [4,2].Desc := 'Secondary Feed Pump', [4,2].RunInterlock := 1, [4,2].OutputAddress := 9, [4,2].InterlockTimer.PRE := 1000, [4,2].InterlockTimer.ACC := 1097, [4,2].InterlockTimer.EN := 1, [4,2].InterlockTimer.DN := 1,
        [4,2].EnableCfg := 1, [4,2].DriveStatus := 1, [4,5].RunOns := 1, [4,5].StopOns := 1, [5,0].InterlockTimer.ACC := 583, [5,0].InterlockTimer.EN := 1, [5,0].InterlockTimer.DN := 1, [5,1].TagName := 'P001', [5,1].Desc := 'Primary Feed Pump', [5,1].RunInterlock := 1, [5,1].OutputAddress := 8, [5,1].InterlockTimer.PRE := 1000, [5,1].InterlockTimer.ACC := 129444, [5,1].InterlockTimer.EN := 1, [5,1].InterlockTimer.DN := 1, [5,1].EnableCfg := 1, [5,1].DriveStatus := 1, [5,2].TagName := 'P002', [5,2].Desc := 'Secondary Feed Pump', [5,2].RunInterlock := 1, [5,2].OutputAddress := 9, [5,2].InterlockTimer.PRE := 1000, [5,2].InterlockTimer.ACC := 129444, [5,2].InterlockTimer.EN := 1, [5,2].InterlockTimer.DN := 1, [5,2].EnableCfg := 1, [5,2].DriveStatus := 1, [5,5].RunOns := 1, [5,5].StopOns := 1);
   ES001 : ALIAS FOR DigitalPoint[2];
   Exchange_OUT : Exchange_OUT;   // Exchange Outputs
   ExternalTCU : BOOL;   // Use of External TCU
   ExternalWeight : BOOL;   // Use of External Weight
   FactorySettings : FactorySettings := (ProductName := 'MTFF80500M3FP1V2/RDP2306026', SerialNumber := 'RDP2306026', ComputerName := 'MTFF80500M3FP1V2', ComputerDesc := 'MTFF80500M3FP1V2_RDP2306026_TFF', DateFormat := 'MM/dd/yyyy', FlagUK := 1, PCV101ClosedSP := 95.0, PCV201ClosedSP := 95.0, TCUDisableSP := 20.0, BagInflateSP := 10.0);
   FI003 : ALIAS FOR AnalogPoint[42];
   FI003Alarm : ALIAS FOR AlarmAnalog[42];
   FI101 : ALIAS FOR AnalogPoint[19];
   FI101_SIG : ALIAS FOR DigitalPoint[110];
   FI101Alarm : ALIAS FOR AlarmAnalog[19];
   FI201 : ALIAS FOR AnalogPoint[2];
   FI201_SIG : ALIAS FOR DigitalPoint[93];
   FI201Alarm : ALIAS FOR AlarmAnalog[2];
   FI401 : ALIAS FOR AnalogPoint[20];
   FI401_SIG : ALIAS FOR DigitalPoint[94];
   FI401Alarm : ALIAS FOR AlarmAnalog[20];
   FirstScanComplete : BOOL := 1;   // First Scan Complete Flag
   FlowPath : FlowPath[64] := ([0].Truth1 := 7168, [0].Mask1 := 7168, [0].Desc := 'Reserved', [1].Status := 1, [1].Truth1 := 387, [1].Mask1 := 2097151, [1].Desc := 'Default', [2].Status := 1, [2].Truth1 := 387, [2].Mask1 := 2097151, [2].Desc := 'Critical', [3].Truth1 := 1114123, [3].Mask1 := 2064527, [3].Desc := 'Single Pass Flush (from inlet manifold)', [4].Truth1 := 1114119, [4].Mask1 := 2064527, [4].Desc := 'Single Pass Flush (from recycle bag)', [5].Truth1 := 1900555, [5].Mask1 := 2064527, [5].Desc := 'System Drain (without recycle bag)', [6].Truth1 := 1900935, [6].Mask1 := 2064783, [6].Desc := 'System Drain (from recycle bag)', [7].Truth1 := 3, [7].Mask1 := 2065283, [7].Desc := 'Membrane Soak', [8].Truth1 := 524928, [8].Mask1 := 2065283, [8].Desc := 'Integrity Test', [9].Truth1 := 768, [9].Mask1 := 2065287, [9].Desc := 'Recycle Bag Fill', [10].Truth1 := 262149, [10].Mask1 := 2065295, [10].Desc := 'Recycle Bag Drain', [11].Truth1 := 131077, [11].Mask1 := 2065295, [11].Desc := 'Recovery Filter Flush', [12].Truth1 := 65927, [12].Mask1 := 2065295, [12].Desc := 'Batch UF or Membrane Recycle', [13].Truth1 := 66439, [13].Mask1 := 2065295, [13].Desc := 'Fed Batch UF or Diafiltration', [14].Truth1 := 131077, [14].Mask1 := 2065295, [14].Desc := 'Product Recovery 1&3  Empty Recycle Bag', [15].Truth1 := 772, [15].Mask1 := 2065295, [15].Desc := 'Product Recovery 2  Empty Retentate Line', [16].Truth1 := 131714, [16].Mask1 := 2065283, [16].Desc := 'Product Recovery 4  Empty membranes', [17].Truth1 := 2065283, [17].Mask1 := 2065283, [17].Desc := 'All Main Flowpath Valves Open', [18].Mask1 := 2065283, [18].Desc := 'All Main Flowpath Valves Closed', [19].Truth1 := 1081355, [19].Mask1 := 2065295,
        [19].Desc := 'Fill Filtrate Line (from inlet manifold)', [20].Truth1 := 33159, [20].Mask1 := 2065295, [20].Desc := 'Fill Filtrate Line (from recycle bag)', [21].Truth1 := 31864, [21].Mask1 := 31868, [21].Desc := 'All Source Valves Open', [22].Status := 1, [22].Mask1 := 31864, [22].Desc := 'All Source Valves Closed', [23].Truth1 := 1024, [23].Mask1 := 31744, [23].Desc := 'Feed Source Open', [24].Truth1 := 2048, [24].Mask1 := 31744, [24].Desc := 'Buffer Source Open', [25].Truth1 := 4096, [25].Mask1 := 31744, [25].Desc := 'Caustic Source Open', [26].Truth1 := 8192, [26].Mask1 := 31744, [26].Desc := 'Water Source Open', [27].Truth1 := 16384, [27].Mask1 := 31744, [27].Desc := 'Air Source Open', [28].Truth1 := 1024, [28].Mask1 := 7168, [28].Desc := 'Feed Source Open - Xfer line', [29].Truth1 := 2048, [29].Mask1 := 7168, [29].Desc := 'Buffer Source Open - Xfer line', [30].Truth1 := 4096, [30].Mask1 := 7168, [30].Desc := 'Air Source Open - Xfer line', [31].Truth1 := 24, [31].Mask1 := 124, [31].Desc := 'Caustic Source Open - Feed line', [32].Truth1 := 40, [32].Mask1 := 124, [32].Desc := 'Water Source Open - Feed line', [33].Truth1 := 72, [33].Mask1 := 124, [33].Desc := 'Buffer/Air Source Open - Feed line', [34].Status := 1, [35].Status := 1, [36].Status := 1, [37].Status := 1, [38].Status := 1, [39].Status := 1, [40].Status := 1, [40].Desc := 'User 1', [41].Status := 1, [41].Desc := 'User 2', [42].Status := 1, [42].Desc := 'User 3', [43].Status := 1, [43].Desc := 'User 4', [44].Status := 1, [44].Desc := 'User 5', [45].Status := 1,
        [46].Status := 1, [47].Status := 1, [48].Status := 1, [49].Status := 1, [50].Status := 1, [51].Status := 1, [52].Status := 1, [53].Status := 1, [54].Status := 1, [55].Status := 1, [56].Status := 1, [57].Status := 1, [58].Status := 1, [59].Status := 1, [60].Status := 1, [61].Truth1 := -1, [61].Mask1 := -1, [62].Mask1 := -1, [63].Status := 1, [63].Truth1 := 387, [63].Mask1 := -1, [63].Mask2 := -1, [63].Mask3 := -1, [63].Mask4 := -1);   // Flow Path Array
        [18]   // All Main Flowpath Valves Closed
        [20]   // Fill Filtrate Line (from recycle bag)
        [10]   // Recycle Bag Drain
        [1]   // Default Flowpath
        [0]   // Reserved : Flowpath Config
        [26]   // Water Source Open
        [11]   // Recovery Filter Flush
        [12]   // Batch UF or Membrane Recycle
        [13]   // Fed Batch UF or Diafiltration
        [14]   // Product Recovery 1&3 – Empty Recycle Bag
        [15]   // Product Recovery 2 – Empty Retentate Line
        [16]   // Product Recovery 4 – Empty membranes
        [17]   // All Main Flowpath Valves Open
        [31]   // Caustic Source Open - Feed line
        [19]   // Fill Filtrate Line (from inlet manifold)
        [9]   // Recycle Bag Fill
        [3]   // Single Pass Flush (from inlet manifold)
        [21]   // All Source Valves Open
        [22]   // All Source Valves Closed
        [23]   // Feed Source Open
        [24]   // Buffer Source Open
        [27]   // Air Source Open
        [28]   // Feed Source Open - Xfer line
        [29]   // Buffer Source Open - Xfer line
        [2]   // Critical Flowpath
        [30]   // Air Source Open - Xfer line
        [32]   // Water Source Open - Feed line
        [33]   // Buffer/Air Source Open - Feed line
        [40]   // User 1
        [41]   // User 2
        [42]   // User 3
        [43]   // User 4
        [44]   // User 5
        [4]   // Single Pass Flush (from recycle bag)
        [5]   // System Drain (without recycle bag)
        [61]   // Reserved : Open All valves
        [62]   // Reserved : Close All valves
        [63]   // Reserved : Saved current flowpath
        [6]   // System Drain (from recycle bag)
        [7]   // Membrane Soak
        [8]   // Integrity Test
        [25]   // Caustic Source Open
   FlowPath_Storage : FlowPath[6,64] := ([0,0].Truth1 := -1, [0,0].Mask1 := -1, [0,0].Desc := 'Reserved', [0,1].Status := 1, [0,1].Truth1 := 539146240, [0,1].Mask1 := -1, [0,1].Desc := 'Default', [0,2].Status := 1, [0,2].Truth1 := 539146240, [0,2].Mask1 := -1, [0,2].Desc := 'Critical', [0,3].Status := 1, [0,3].Mask1 := 2047, [0,3].Desc := 'Close All Inlets', [0,4].Truth1 := 17, [0,4].Mask1 := 63, [0,4].Desc := 'Inlet 1A', [0,5].Truth1 := 18, [0,5].Mask1 := 63, [0,5].Desc := 'Inlet 1B', [0,6].Truth1 := 20, [0,6].Mask1 := 63, [0,6].Desc := 'Inlet 1C', [0,7].Truth1 := 24, [0,7].Mask1 := 63, [0,7].Desc := 'Inlet 1D', [0,8].Truth1 := 32, [0,8].Mask1 := 63, [0,8].Desc := 'Inlet 1E', [0,9].Truth1 := 64, [0,9].Mask1 := 1984, [0,9].Desc := 'Inlet 2A', [0,10].Truth1 := 128, [0,10].Mask1 := 1984, [0,10].Desc := 'Inlet 2B', [0,11].Truth1 := 256, [0,11].Mask1 := 1984, [0,11].Desc := 'Inlet 2C', [0,12].Truth1 := 512, [0,12].Mask1 := 1984, [0,12].Desc := 'Inlet 2D', [0,13].Truth1 := 1024, [0,13].Mask1 := 1984, [0,13].Desc := 'Inlet 2E', [0,14].Truth1 := 2047, [0,14].Mask1 := 2047, [0,14].Desc := 'Open All Inlets', [0,15].Truth1 := 2047, [0,15].Mask1 := 2047, [0,15].Desc := 'Flexware Installation', [0,16].Truth1 := 2048, [0,16].Mask1 := -2147477504, [0,16].Desc := 'P001 Process', [0,17].Truth1 := -2147481600, [0,17].Mask1 := -2147477504, [0,17].Desc := 'P001 Drain', [0,18].Truth1 := 4096, [0,18].Mask1 := -2147477504, [0,18].Desc := 'P002 Process', [0,19].Truth1 := -2147479552,
        [0,19].Mask1 := -2147477504, [0,19].Desc := 'P002 Drain', [0,20].Status := 1, [0,20].Truth1 := 6144, [0,20].Mask1 := -2147477504, [0,20].Desc := 'Dual Pumps Process', [0,21].Truth1 := -2147477504, [0,21].Mask1 := -2147477504, [0,21].Desc := 'Dual Pumps Drain', [0,22].Status := 1, [0,22].Truth1 := 40960, [0,22].Mask1 := -1073684480, [0,22].Desc := 'BBT Online', [0,23].Truth1 := 16384, [0,23].Mask1 := -1073684480, [0,23].Desc := 'BBT Bypass', [0,24].Truth1 := 1073741824, [0,24].Mask1 := 1073741824, [0,24].Desc := 'BBT Vent', [0,25].Truth1 := 1073750016, [0,25].Mask1 := -1073684480, [0,25].Desc := 'BBT Clean', [0,26].Truth1 := -1073692672, [0,26].Mask1 := -1073684480, [0,26].Desc := 'BBT Drain', [0,27].Mask1 := -1, [0,27].Desc := 'BBT User', [0,28].Truth1 := 327680, [0,28].Mask1 := 458752, [0,28].Desc := 'Filter Online', [0,29].Status := 1, [0,29].Truth1 := 131072, [0,29].Mask1 := 458752, [0,29].Desc := 'Filter Bypass', [0,30].Mask1 := -1, [0,30].Desc := 'Filter User', [0,31].Truth1 := 59244544, [0,31].Mask1 := 66584576, [0,31].Desc := 'Column Forward', [0,32].Truth1 := 55574528, [0,32].Mask1 := 66584576, [0,32].Desc := 'Column Reverse', [0,33].Status := 1, [0,33].Truth1 := 2097152, [0,33].Mask1 := 66584576, [0,33].Desc := 'Column Bypass', [0,34].Mask1 := -1, [0,34].Desc := 'Column user', [0,35].Status := 1, [0,35].Truth1 := 536870912, [0,35].Mask1 := 1006632960, [0,35].Desc := 'Fraction Waste', [0,36].Truth1 := 268435456, [0,36].Mask1 := 1006632960, [0,36].Desc := 'Fraction 3', [0,37].Truth1 := 134217728, [0,37].Mask1 := 1006632960, [0,37].Desc := 'Fraction 2', [0,38].Truth1 := 67108864, [0,38].Mask1 := 1006632960,
        [0,38].Desc := 'Fraction 1', [0,39].Truth1 := -1, [0,39].Mask1 := -1, [0,39].Desc := 'System Drain', [0,40].Status := 1, [0,40].Desc := 'User 1', [0,41].Status := 1, [0,41].Desc := 'User 2', [0,42].Truth2 := 32768, [0,42].Mask2 := 32960, [0,42].Desc := 'User 3', [0,43].Status := 1, [0,43].Desc := 'User 4', [0,44].Truth1 := 118489088, [0,44].Mask1 := 133169152, [0,44].Desc := 'User 5', [0,45].Status := 1, [0,46].Status := 1, [0,47].Status := 1, [0,48].Status := 1, [0,49].Status := 1, [0,50].Status := 1, [0,51].Status := 1, [0,52].Status := 1, [0,53].Status := 1, [0,54].Status := 1, [0,55].Status := 1, [0,56].Status := 1, [0,57].Status := 1, [0,58].Status := 1, [0,59].Status := 1, [0,60].Status := 1, [0,61].Truth1 := -1, [0,61].Mask1 := -1, [0,62].Mask1 := -1, [0,63].Status := 1, [0,63].Truth1 := 539146240, [0,63].Mask1 := -1, [0,63].Mask2 := -1, [0,63].Mask3 := -1, [0,63].Mask4 := -1, [1,0].Truth1 := -1, [1,0].Mask1 := -1, [1,0].Desc := 'Reserved', [1,1].Status := 1, [1,1].Truth1 := 539146240, [1,1].Mask1 := -1, [1,1].Desc := 'Default', [1,2].Status := 1, [1,2].Truth1 := 539146240, [1,2].Mask1 := -1, [1,2].Desc := 'Critical', [1,3].Status := 1, [1,3].Mask1 := 2047, [1,3].Desc := 'Close All Inlets', [1,4].Truth1 := 17, [1,4].Mask1 := 63, [1,4].Desc := 'Inlet 1A', [1,5].Truth1 := 18, [1,5].Mask1 := 63,
        [1,5].Desc := 'Inlet 1B', [1,6].Truth1 := 20, [1,6].Mask1 := 63, [1,6].Desc := 'Inlet 1C', [1,7].Truth1 := 24, [1,7].Mask1 := 63, [1,7].Desc := 'Inlet 1D', [1,8].Truth1 := 32, [1,8].Mask1 := 63, [1,8].Desc := 'Inlet 1E', [1,9].Truth1 := 64, [1,9].Mask1 := 1984, [1,9].Desc := 'Inlet 2A', [1,10].Truth1 := 128, [1,10].Mask1 := 1984, [1,10].Desc := 'Inlet 2B', [1,11].Truth1 := 256, [1,11].Mask1 := 1984, [1,11].Desc := 'Inlet 2C', [1,12].Truth1 := 512, [1,12].Mask1 := 1984, [1,12].Desc := 'Inlet 2D', [1,13].Truth1 := 1024, [1,13].Mask1 := 1984, [1,13].Desc := 'Inlet 2E', [1,14].Truth1 := 2047, [1,14].Mask1 := 2047, [1,14].Desc := 'Open All Inlets', [1,15].Truth1 := 2047, [1,15].Mask1 := 2047, [1,15].Desc := 'Flexware Installation', [1,16].Truth1 := 2048, [1,16].Mask1 := -2147477504, [1,16].Desc := 'P001 Process', [1,17].Truth1 := -2147481600, [1,17].Mask1 := -2147477504, [1,17].Desc := 'P001 Drain', [1,18].Truth1 := 4096, [1,18].Mask1 := -2147477504, [1,18].Desc := 'P002 Process', [1,19].Truth1 := -2147479552, [1,19].Mask1 := -2147477504, [1,19].Desc := 'P002 Drain', [1,20].Status := 1, [1,20].Truth1 := 6144, [1,20].Mask1 := -2147477504, [1,20].Desc := 'Dual Pumps Process', [1,21].Truth1 := -2147477504, [1,21].Mask1 := -2147477504, [1,21].Desc := 'Dual Pumps Drain', [1,22].Status := 1, [1,22].Truth1 := 40960, [1,22].Mask1 := -1073684480, [1,22].Desc := 'BBT Online', [1,23].Truth1 := 16384, [1,23].Mask1 := -1073684480, [1,23].Desc := 'BBT Bypass', [1,24].Truth1 := 1073741824, [1,24].Mask1 := 1073741824, [1,24].Desc := 'BBT Vent',
        [1,25].Truth1 := 1073750016, [1,25].Mask1 := -1073684480, [1,25].Desc := 'BBT Clean', [1,26].Truth1 := -1073692672, [1,26].Mask1 := -1073684480, [1,26].Desc := 'BBT Drain', [1,27].Mask1 := -1, [1,27].Desc := 'BBT User', [1,28].Truth1 := 327680, [1,28].Mask1 := 458752, [1,28].Desc := 'Filter Online', [1,29].Status := 1, [1,29].Truth1 := 131072, [1,29].Mask1 := 458752, [1,29].Desc := 'Filter Bypass', [1,30].Mask1 := -1, [1,30].Desc := 'Filter User', [1,31].Truth1 := 59244544, [1,31].Mask1 := 66584576, [1,31].Desc := 'Column Forward', [1,32].Truth1 := 55574528, [1,32].Mask1 := 66584576, [1,32].Desc := 'Column Reverse', [1,33].Status := 1, [1,33].Truth1 := 2097152, [1,33].Mask1 := 66584576, [1,33].Desc := 'Column Bypass', [1,34].Mask1 := -1, [1,34].Desc := 'Column user', [1,35].Status := 1, [1,35].Truth1 := 536870912, [1,35].Mask1 := 1006632960, [1,35].Desc := 'Fraction Waste', [1,36].Truth1 := 268435456, [1,36].Mask1 := 1006632960, [1,36].Desc := 'Fraction 3', [1,37].Truth1 := 134217728, [1,37].Mask1 := 1006632960, [1,37].Desc := 'Fraction 2', [1,38].Truth1 := 67108864, [1,38].Mask1 := 1006632960, [1,38].Desc := 'Fraction 1', [1,39].Truth1 := -1, [1,39].Mask1 := -1, [1,39].Desc := 'System Drain', [1,40].Status := 1, [1,40].Desc := 'User 1', [1,41].Status := 1, [1,41].Desc := 'User 2', [1,42].Truth2 := 32768, [1,42].Mask2 := 32960, [1,42].Desc := 'User 3', [1,43].Status := 1, [1,43].Desc := 'User 4', [1,44].Truth1 := 118489088, [1,44].Mask1 := 133169152, [1,44].Desc := 'User 5', [1,45].Status := 1, [1,46].Status := 1, [1,47].Status := 1,
        [1,48].Status := 1, [1,49].Status := 1, [1,50].Status := 1, [1,51].Status := 1, [1,52].Status := 1, [1,53].Status := 1, [1,54].Status := 1, [1,55].Status := 1, [1,56].Status := 1, [1,57].Status := 1, [1,58].Status := 1, [1,59].Status := 1, [1,60].Status := 1, [1,61].Truth1 := -1, [1,61].Mask1 := -1, [1,62].Mask1 := -1, [1,63].Status := 1, [1,63].Truth1 := 539146240, [1,63].Mask1 := -1, [1,63].Mask2 := -1, [1,63].Mask3 := -1, [1,63].Mask4 := -1, [2,0].Truth1 := -1, [2,0].Mask1 := -1, [2,0].Desc := 'Reserved', [2,1].Status := 1, [2,1].Truth1 := 539146240, [2,1].Mask1 := -1, [2,1].Desc := 'Default', [2,2].Status := 1, [2,2].Truth1 := 539146240, [2,2].Mask1 := -1, [2,2].Desc := 'Critical', [2,3].Status := 1, [2,3].Mask1 := 2047, [2,3].Desc := 'Close All Inlets', [2,4].Truth1 := 17, [2,4].Mask1 := 63, [2,4].Desc := 'Inlet 1A', [2,5].Truth1 := 18, [2,5].Mask1 := 63, [2,5].Desc := 'Inlet 1B', [2,6].Truth1 := 20, [2,6].Mask1 := 63, [2,6].Desc := 'Inlet 1C', [2,7].Truth1 := 24, [2,7].Mask1 := 63, [2,7].Desc := 'Inlet 1D', [2,8].Truth1 := 32, [2,8].Mask1 := 63, [2,8].Desc := 'Inlet 1E', [2,9].Truth1 := 64, [2,9].Mask1 := 1984, [2,9].Desc := 'Inlet 2A', [2,10].Truth1 := 128, [2,10].Mask1 := 1984, [2,10].Desc := 'Inlet 2B', [2,11].Truth1 := 256, [2,11].Mask1 := 1984, [2,11].Desc := 'Inlet 2C',
        [2,12].Truth1 := 512, [2,12].Mask1 := 1984, [2,12].Desc := 'Inlet 2D', [2,13].Truth1 := 1024, [2,13].Mask1 := 1984, [2,13].Desc := 'Inlet 2E', [2,14].Truth1 := 2047, [2,14].Mask1 := 2047, [2,14].Desc := 'Open All Inlets', [2,15].Truth1 := 2047, [2,15].Mask1 := 2047, [2,15].Desc := 'Flexware Installation', [2,16].Truth1 := 2048, [2,16].Mask1 := -2147477504, [2,16].Desc := 'P001 Process', [2,17].Truth1 := -2147481600, [2,17].Mask1 := -2147477504, [2,17].Desc := 'P001 Drain', [2,18].Truth1 := 4096, [2,18].Mask1 := -2147477504, [2,18].Desc := 'P002 Process', [2,19].Truth1 := -2147479552, [2,19].Mask1 := -2147477504, [2,19].Desc := 'P002 Drain', [2,20].Status := 1, [2,20].Truth1 := 6144, [2,20].Mask1 := -2147477504, [2,20].Desc := 'Dual Pumps Process', [2,21].Truth1 := -2147477504, [2,21].Mask1 := -2147477504, [2,21].Desc := 'Dual Pumps Drain', [2,22].Status := 1, [2,22].Truth1 := 40960, [2,22].Mask1 := -1073684480, [2,22].Desc := 'BBT Online', [2,23].Truth1 := 16384, [2,23].Mask1 := -1073684480, [2,23].Desc := 'BBT Bypass', [2,24].Truth1 := 1073741824, [2,24].Mask1 := 1073741824, [2,24].Desc := 'BBT Vent', [2,25].Truth1 := 1073750016, [2,25].Mask1 := -1073684480, [2,25].Desc := 'BBT Clean', [2,26].Truth1 := -1073692672, [2,26].Mask1 := -1073684480, [2,26].Desc := 'BBT Drain', [2,27].Mask1 := -1, [2,27].Desc := 'BBT User', [2,28].Truth1 := 327680, [2,28].Mask1 := 458752, [2,28].Desc := 'Filter Online', [2,29].Status := 1, [2,29].Truth1 := 131072, [2,29].Mask1 := 458752, [2,29].Desc := 'Filter Bypass', [2,30].Mask1 := -1, [2,30].Desc := 'Filter User', [2,31].Truth1 := 59244544, [2,31].Mask1 := 66584576,
        [2,31].Desc := 'Column Forward', [2,32].Truth1 := 55574528, [2,32].Mask1 := 66584576, [2,32].Desc := 'Column Reverse', [2,33].Status := 1, [2,33].Truth1 := 2097152, [2,33].Mask1 := 66584576, [2,33].Desc := 'Column Bypass', [2,34].Mask1 := -1, [2,34].Desc := 'Column user', [2,35].Status := 1, [2,35].Truth1 := 536870912, [2,35].Mask1 := 1006632960, [2,35].Desc := 'Fraction Waste', [2,36].Truth1 := 268435456, [2,36].Mask1 := 1006632960, [2,36].Desc := 'Fraction 3', [2,37].Truth1 := 134217728, [2,37].Mask1 := 1006632960, [2,37].Desc := 'Fraction 2', [2,38].Truth1 := 67108864, [2,38].Mask1 := 1006632960, [2,38].Desc := 'Fraction 1', [2,39].Truth1 := -1, [2,39].Mask1 := -1, [2,39].Desc := 'System Drain', [2,40].Status := 1, [2,40].Desc := 'User 1', [2,41].Status := 1, [2,41].Desc := 'User 2', [2,42].Truth2 := 32768, [2,42].Mask2 := 32960, [2,42].Desc := 'User 3', [2,43].Status := 1, [2,43].Desc := 'User 4', [2,44].Truth1 := 118489088, [2,44].Mask1 := 133169152, [2,44].Desc := 'User 5', [2,45].Status := 1, [2,46].Status := 1, [2,47].Status := 1, [2,48].Status := 1, [2,49].Status := 1, [2,50].Status := 1, [2,51].Status := 1, [2,52].Status := 1, [2,53].Status := 1, [2,54].Status := 1, [2,55].Status := 1, [2,56].Status := 1, [2,57].Status := 1, [2,58].Status := 1, [2,59].Status := 1, [2,60].Status := 1, [2,61].Truth1 := -1, [2,61].Mask1 := -1, [2,62].Mask1 := -1, [2,63].Status := 1, [2,63].Truth1 := 539146240, [2,63].Mask1 := -1,
        [2,63].Mask2 := -1, [2,63].Mask3 := -1, [2,63].Mask4 := -1, [3,0].Status := 1, [3,1].Status := 1, [3,2].Truth1 := 539146240, [3,2].Mask1 := -1, [3,3].Status := 1, [3,3].Mask1 := 2047, [3,4].Truth1 := 17, [3,4].Mask1 := 63, [3,5].Truth1 := 18, [3,5].Mask1 := 63, [3,6].Truth1 := 20, [3,6].Mask1 := 63, [3,7].Truth1 := 24, [3,7].Mask1 := 63, [3,8].Truth1 := 32, [3,8].Mask1 := 63, [3,9].Truth1 := 64, [3,9].Mask1 := 1984, [3,10].Truth1 := 128, [3,10].Mask1 := 1984, [3,11].Truth1 := 256, [3,11].Mask1 := 1984, [3,12].Truth1 := 512, [3,12].Mask1 := 1984, [3,13].Truth1 := 1024, [3,13].Mask1 := 1984, [3,14].Truth1 := 2047, [3,14].Mask1 := 2047, [3,15].Truth1 := 2047, [3,15].Mask1 := 2047, [3,16].Truth1 := 2048, [3,16].Mask1 := -2147477504, [3,17].Truth1 := -2147481600, [3,17].Mask1 := -2147477504, [3,18].Truth1 := 4096, [3,18].Mask1 := -2147477504, [3,19].Truth1 := -2147479552, [3,19].Mask1 := -2147477504, [3,20].Truth1 := 6144, [3,20].Mask1 := -2147477504, [3,21].Truth1 := -2147477504, [3,21].Mask1 := -2147477504, [3,22].Truth1 := 40960, [3,22].Mask1 := -1073684480, [3,23].Truth1 := 16384, [3,23].Mask1 := -1073684480, [3,24].Truth1 := 1073741824, [3,24].Mask1 := 1073741824, [3,25].Truth1 := 1073750016, [3,25].Mask1 := -1073684480, [3,26].Truth1 := -1073692672, [3,26].Mask1 := -1073684480, [3,27].Status := 1, [3,28].Truth1 := 327680, [3,28].Mask1 := 458752, [3,29].Truth1 := 131072, [3,29].Mask1 := 458752,
        [3,30].Status := 1, [3,31].Truth1 := 59244544, [3,31].Mask1 := 66584576, [3,32].Truth1 := 55574528, [3,32].Mask1 := 66584576, [3,33].Truth1 := 2097152, [3,33].Mask1 := 66584576, [3,34].Status := 1, [3,35].Truth1 := 536870912, [3,35].Mask1 := 1006632960, [3,36].Truth1 := 268435456, [3,36].Mask1 := 1006632960, [3,37].Truth1 := 134217728, [3,37].Mask1 := 1006632960, [3,38].Truth1 := 67108864, [3,38].Mask1 := 1006632960, [3,39].Truth1 := -1, [3,39].Mask1 := -1, [3,40].Status := 1, [3,41].Status := 1, [3,42].Status := 1, [3,43].Status := 1, [3,44].Status := 1, [3,45].Status := 1, [3,46].Status := 1, [3,47].Status := 1, [3,48].Status := 1, [3,49].Status := 1, [3,50].Status := 1, [3,51].Status := 1, [3,52].Status := 1, [3,53].Status := 1, [3,54].Status := 1, [3,55].Status := 1, [3,56].Status := 1, [3,57].Status := 1, [3,58].Status := 1, [3,59].Status := 1, [3,60].Status := 1, [3,61].Truth1 := -1, [3,61].Mask1 := -1, [3,62].Status := 1, [3,62].Mask1 := -1, [3,63].Status := 1, [4,0].Truth1 := -1, [4,0].Mask1 := -1, [4,0].Desc := 'Reserved', [4,1].Status := 1, [4,1].Truth1 := 539146240, [4,1].Mask1 := -1, [4,1].Desc := 'Default', [4,2].Status := 1, [4,2].Truth1 := 539146240, [4,2].Mask1 := -1, [4,2].Desc := 'Critical', [4,3].Status := 1, [4,3].Mask1 := 2047, [4,3].Desc := 'Close All Inlets', [4,4].Truth1 := 17, [4,4].Mask1 := 63,
        [4,4].Desc := 'Inlet 1A', [4,5].Truth1 := 18, [4,5].Mask1 := 63, [4,5].Desc := 'Inlet 1B', [4,6].Truth1 := 20, [4,6].Mask1 := 63, [4,6].Desc := 'Inlet 1C', [4,7].Truth1 := 24, [4,7].Mask1 := 63, [4,7].Desc := 'Inlet 1D', [4,8].Truth1 := 32, [4,8].Mask1 := 63, [4,8].Desc := 'Inlet 1E', [4,9].Truth1 := 64, [4,9].Mask1 := 1984, [4,9].Desc := 'Inlet 2A', [4,10].Truth1 := 128, [4,10].Mask1 := 1984, [4,10].Desc := 'Inlet 2B', [4,11].Truth1 := 256, [4,11].Mask1 := 1984, [4,11].Desc := 'Inlet 2C', [4,12].Truth1 := 512, [4,12].Mask1 := 1984, [4,12].Desc := 'Inlet 2D', [4,13].Truth1 := 1024, [4,13].Mask1 := 1984, [4,13].Desc := 'Inlet 2E', [4,14].Truth1 := 2047, [4,14].Mask1 := 2047, [4,14].Desc := 'Open All Inlets', [4,15].Truth1 := 2047, [4,15].Mask1 := 2047, [4,15].Desc := 'Flexware Installation', [4,16].Truth1 := 4096, [4,16].Mask1 := -2147477504, [4,16].Desc := 'P001 Process', [4,17].Truth1 := -2147479552, [4,17].Mask1 := -2147477504, [4,17].Desc := 'P001 Drain', [4,18].Truth1 := 2048, [4,18].Mask1 := -2147477504, [4,18].Desc := 'P002 Process', [4,19].Truth1 := -2147481600, [4,19].Mask1 := -2147477504, [4,19].Desc := 'P002 Drain', [4,20].Status := 1, [4,20].Truth1 := 6144, [4,20].Mask1 := -2147477504, [4,20].Desc := 'Dual Pumps Process', [4,21].Truth1 := -2147477504, [4,21].Mask1 := -2147477504, [4,21].Desc := 'Dual Pumps Drain', [4,22].Status := 1, [4,22].Truth1 := 40960, [4,22].Mask1 := -1073684480, [4,22].Desc := 'BBT Online', [4,23].Truth1 := 16384, [4,23].Mask1 := -1073684480, [4,23].Desc := 'BBT Bypass',
        [4,24].Truth1 := 1073741824, [4,24].Mask1 := 1073741824, [4,24].Desc := 'BBT Vent', [4,25].Truth1 := 1073750016, [4,25].Mask1 := -1073684480, [4,25].Desc := 'BBT Clean', [4,26].Truth1 := -1073692672, [4,26].Mask1 := -1073684480, [4,26].Desc := 'BBT Drain', [4,27].Mask1 := -1, [4,27].Desc := 'BBT User', [4,28].Truth1 := 327680, [4,28].Mask1 := 458752, [4,28].Desc := 'Filter Online', [4,29].Status := 1, [4,29].Truth1 := 131072, [4,29].Mask1 := 458752, [4,29].Desc := 'Filter Bypass', [4,30].Mask1 := -1, [4,30].Desc := 'Filter User', [4,31].Truth1 := 59244544, [4,31].Mask1 := 66584576, [4,31].Desc := 'Column Forward', [4,32].Truth1 := 55574528, [4,32].Mask1 := 66584576, [4,32].Desc := 'Column Reverse', [4,33].Status := 1, [4,33].Truth1 := 2097152, [4,33].Mask1 := 66584576, [4,33].Desc := 'Column Bypass', [4,34].Mask1 := -1, [4,34].Desc := 'Column user', [4,35].Status := 1, [4,35].Truth1 := 536870912, [4,35].Mask1 := 1006632960, [4,35].Desc := 'Fraction Waste', [4,36].Truth1 := 268435456, [4,36].Mask1 := 1006632960, [4,36].Desc := 'Fraction 3', [4,37].Truth1 := 134217728, [4,37].Mask1 := 1006632960, [4,37].Desc := 'Fraction 2', [4,38].Truth1 := 67108864, [4,38].Mask1 := 1006632960, [4,38].Desc := 'Fraction 1', [4,39].Truth1 := -1, [4,39].Mask1 := -1, [4,39].Desc := 'System Drain', [4,40].Status := 1, [4,40].Desc := 'User 1', [4,41].Status := 1, [4,41].Desc := 'User 2', [4,42].Truth2 := 32768, [4,42].Mask2 := 32960, [4,42].Desc := 'User 3', [4,43].Status := 1, [4,43].Desc := 'User 4', [4,44].Truth1 := 118489088, [4,44].Mask1 := 133169152, [4,44].Desc := 'User 5',
        [4,45].Status := 1, [4,46].Status := 1, [4,47].Status := 1, [4,48].Status := 1, [4,49].Status := 1, [4,50].Status := 1, [4,51].Status := 1, [4,52].Status := 1, [4,53].Status := 1, [4,54].Status := 1, [4,55].Status := 1, [4,56].Status := 1, [4,57].Status := 1, [4,58].Status := 1, [4,59].Status := 1, [4,60].Status := 1, [4,61].Truth1 := -1, [4,61].Mask1 := -1, [4,62].Mask1 := -1, [4,63].Status := 1, [4,63].Truth1 := 539146240, [4,63].Mask1 := -1, [4,63].Mask2 := -1, [4,63].Mask3 := -1, [4,63].Mask4 := -1, [5,0].Truth1 := -1, [5,0].Mask1 := -1, [5,0].Desc := 'Reserved', [5,1].Status := 1, [5,1].Truth1 := 539146240, [5,1].Mask1 := -1, [5,1].Desc := 'Default', [5,2].Status := 1, [5,2].Truth1 := 539146240, [5,2].Mask1 := -1, [5,2].Desc := 'Critical', [5,3].Status := 1, [5,3].Mask1 := 2047, [5,3].Desc := 'Close All Inlets', [5,4].Truth1 := 17, [5,4].Mask1 := 63, [5,4].Desc := 'Inlet 1A', [5,5].Truth1 := 18, [5,5].Mask1 := 63, [5,5].Desc := 'Inlet 1B', [5,6].Truth1 := 20, [5,6].Mask1 := 63, [5,6].Desc := 'Inlet 1C', [5,7].Truth1 := 24, [5,7].Mask1 := 63, [5,7].Desc := 'Inlet 1D', [5,8].Truth1 := 32, [5,8].Mask1 := 63, [5,8].Desc := 'Inlet 1E', [5,9].Truth1 := 64, [5,9].Mask1 := 1984, [5,9].Desc := 'Inlet 2A', [5,10].Truth1 := 128, [5,10].Mask1 := 1984, [5,10].Desc := 'Inlet 2B',
        [5,11].Truth1 := 256, [5,11].Mask1 := 1984, [5,11].Desc := 'Inlet 2C', [5,12].Truth1 := 512, [5,12].Mask1 := 1984, [5,12].Desc := 'Inlet 2D', [5,13].Truth1 := 1024, [5,13].Mask1 := 1984, [5,13].Desc := 'Inlet 2E', [5,14].Truth1 := 2047, [5,14].Mask1 := 2047, [5,14].Desc := 'Open All Inlets', [5,15].Truth1 := 2047, [5,15].Mask1 := 2047, [5,15].Desc := 'Flexware Installation', [5,16].Truth1 := 2048, [5,16].Mask1 := -2147477504, [5,16].Desc := 'P001 Process', [5,17].Truth1 := -2147481600, [5,17].Mask1 := -2147477504, [5,17].Desc := 'P001 Drain', [5,18].Truth1 := 4096, [5,18].Mask1 := -2147477504, [5,18].Desc := 'P002 Process', [5,19].Truth1 := -2147479552, [5,19].Mask1 := -2147477504, [5,19].Desc := 'P002 Drain', [5,20].Status := 1, [5,20].Truth1 := 6144, [5,20].Mask1 := -2147477504, [5,20].Desc := 'Dual Pumps Process', [5,21].Truth1 := -2147477504, [5,21].Mask1 := -2147477504, [5,21].Desc := 'Dual Pumps Drain', [5,22].Status := 1, [5,22].Truth1 := 40960, [5,22].Mask1 := -1073684480, [5,22].Desc := 'BBT Online', [5,23].Truth1 := 16384, [5,23].Mask1 := -1073684480, [5,23].Desc := 'BBT Bypass', [5,24].Truth1 := 1073741824, [5,24].Mask1 := 1073741824, [5,24].Desc := 'BBT Vent', [5,25].Truth1 := 1073750016, [5,25].Mask1 := -1073684480, [5,25].Desc := 'BBT Clean', [5,26].Truth1 := -1073692672, [5,26].Mask1 := -1073684480, [5,26].Desc := 'BBT Drain', [5,27].Mask1 := -1, [5,27].Desc := 'BBT User', [5,28].Truth1 := 327680, [5,28].Mask1 := 458752, [5,28].Desc := 'Filter Online', [5,29].Status := 1, [5,29].Truth1 := 131072, [5,29].Mask1 := 458752, [5,29].Desc := 'Filter Bypass', [5,30].Mask1 := -1,
        [5,30].Desc := 'Filter User', [5,31].Truth1 := 59244544, [5,31].Mask1 := 66584576, [5,31].Desc := 'Column Forward', [5,32].Truth1 := 55574528, [5,32].Mask1 := 66584576, [5,32].Desc := 'Column Reverse', [5,33].Status := 1, [5,33].Truth1 := 2097152, [5,33].Mask1 := 66584576, [5,33].Desc := 'Column Bypass', [5,34].Mask1 := -1, [5,34].Desc := 'Column user', [5,35].Status := 1, [5,35].Truth1 := 536870912, [5,35].Mask1 := 1006632960, [5,35].Desc := 'Fraction Waste', [5,36].Truth1 := 268435456, [5,36].Mask1 := 1006632960, [5,36].Desc := 'Fraction 3', [5,37].Truth1 := 134217728, [5,37].Mask1 := 1006632960, [5,37].Desc := 'Fraction 2', [5,38].Truth1 := 67108864, [5,38].Mask1 := 1006632960, [5,38].Desc := 'Fraction 1', [5,39].Truth1 := -1, [5,39].Mask1 := -1, [5,39].Desc := 'System Drain', [5,40].Status := 1, [5,40].Desc := 'User 1', [5,41].Status := 1, [5,41].Desc := 'User 2', [5,42].Truth2 := 32768, [5,42].Mask2 := 32960, [5,42].Desc := 'User 3', [5,43].Status := 1, [5,43].Desc := 'User 4', [5,44].Truth1 := 118489088, [5,44].Mask1 := 133169152, [5,44].Desc := 'User 5', [5,45].Status := 1, [5,46].Status := 1, [5,47].Status := 1, [5,48].Status := 1, [5,49].Status := 1, [5,50].Status := 1, [5,51].Status := 1, [5,52].Status := 1, [5,53].Status := 1, [5,54].Status := 1, [5,55].Status := 1, [5,56].Status := 1, [5,57].Status := 1, [5,58].Status := 1, [5,59].Status := 1, [5,60].Status := 1, [5,61].Truth1 := -1, [5,61].Mask1 := -1, [5,62].Mask1 := -1,
        [5,63].Status := 1, [5,63].Truth1 := 539146240, [5,63].Mask1 := -1, [5,63].Mask2 := -1, [5,63].Mask3 := -1, [5,63].Mask4 := -1);
   FlowPathControl : FlowPathControl := (Valve1 := 387, MaxFlowPath := 63, Status := 63, StatusHMI := 63, Save := 1, SaveOns := 1, FlowpathEnable[0] := 1, FlowpathEnable[1] := 1, FlowpathEnable[2] := 1, FlowpathEnable[3] := 1, FlowpathEnable[4] := 1, FlowpathEnable[5] := 1, FlowpathEnable[6] := 1, FlowpathEnable[7] := 1, FlowpathEnable[8] := 1, FlowpathEnable[9] := 1, FlowpathEnable[10] := 1, FlowpathEnable[11] := 1, FlowpathEnable[12] := 1, FlowpathEnable[13] := 1, FlowpathEnable[14] := 1, FlowpathEnable[15] := 1, FlowpathEnable[16] := 1, FlowpathEnable[17] := 1, FlowpathEnable[18] := 1, FlowpathEnable[19] := 1, FlowpathEnable[20] := 1, FlowpathEnable[21] := 1, FlowpathEnable[22] := 1, FlowpathEnable[23] := 1, FlowpathEnable[24] := 1, FlowpathEnable[25] := 1, FlowpathEnable[26] := 1, FlowpathEnable[27] := 1, FlowpathEnable[28] := 1, FlowpathEnable[29] := 1, FlowpathEnable[30] := 1, FlowpathEnable[31] := 1, FlowpathEnable[32] := 1, FlowpathEnable[33] := 1, FlowpathEnable[34] := 1, FlowpathEnable[35] := 1, FlowpathEnable[36] := 1, FlowpathEnable[37] := 1, FlowpathEnable[38] := 1, FlowpathEnable[39] := 1, FlowpathEnable[40] := 1, FlowpathEnable[41] := 1, FlowpathEnable[42] := 1, FlowpathEnable[43] := 1, FlowpathEnable[44] := 1, FlowpathEnable[45] := 1, FlowpathEnable[46] := 1, FlowpathEnable[47] := 1, FlowpathEnable[48] := 1, FlowpathEnable[49] := 1, FlowpathEnable[50] := 1, FlowpathEnable[51] := 1, FlowpathEnable[52] := 1, FlowpathEnable[53] := 1,
        FlowpathEnable[54] := 1, FlowpathEnable[55] := 1, FlowpathEnable[56] := 1, FlowpathEnable[57] := 1, FlowpathEnable[58] := 1, FlowpathEnable[59] := 1, FlowpathEnable[60] := 1, FlowpathEnable[61] := 1, FlowpathEnable[62] := 1, FlowpathEnable[63] := 1, SaveStored := 1, HoldOns := 1);   // Flow Path Control
   FlowPathSetup : FlowPathSetup := (Number := 1, Prev := 1);   // Flow Path Setup Data
   FQ_Conc : ALIAS FOR Totalizer[0];   // Concentration Totalizer
   FQ_Diaf : ALIAS FOR Totalizer[1];   // DiafiltrationTotalizer
   Gateway : Gateway := (Inhibition := 4, Input[22] := 5856, Input[23] := 5856, Output[1] := 54984, Output[2] := 110041, Output[3] := 8212, Output[4] := 25729, Output[5] := -41, Output[6] := -25, Output[7] := -99, Output[8] := 7560, Output[9] := -94, Output[11] := 20, Output[13] := 18, Output[15] := -500, Output[16] := -500, Output[17] := -2500, Output[18] := -2500, Output[19] := -2500, Output[20] := -24997, Output[21] := -24997, Output[28] := 21878, Output[29] := 21878, Output[30] := 21878, Output[31] := 21878, Output[46] := 100000, Output[50] := -25000, Output[56] := 65994807, Output[57] := 1352834048, Output[58] := 1715480648, Output[59] := 23579, Output[64] := 10312, Output[82] := 1, Output[106] := 5866, Output[107] := 5856, Watchdog_Heartbeat_Timer.TimerEnable := 1, Watchdog_Heartbeat_Timer.ACC := 89, Watchdog_Heartbeat_Timer.EN := 1, Watchdog_Heartbeat_Timer.DN := 1, Watchdog_In_Ext := 5856, Watchdog_In_Skid := 5856, Watchdog_Out_Ext := 5856, Watchdog_Out_Skid := 5866, Index := 64, Index2 := 32);   // Gateway Control
   GradientLinear : LinearGradient := (Variable := 1, Basis := 1, Y[0] := 50.0);   // (To be keep to avoid error on Recipe Download)
   GWModbus : IO_Station := (Node_Comm_Status_value := 12288);   // Status of Gateway Modbus
   HoldTime : ALIAS FOR Timers[20];   // Hold Time
   HTCCollectorError : BOOL;   // Historical Data Collector Error (Set to 1 by HMI if Error)
   HTCHeartBeat : BOOL;   // Historical Data Collection heartbeat (Set to 1 by HMI Reset to 0 by PLC)
   IBA001 : ALIAS FOR DigitalOutput[25];
   LI101 : ALIAS FOR AnalogPoint[44];
   LI101Alarm : ALIAS FOR AlarmAnalog[44];
   LogVal : LoggedValue;   // Setpoints to be logged
        .Value[0]   // P001 Manual setpoint
        .Value[1]   // P001 Flow setpoint
        .Value[2]   // P001 Linear Velocity setpoint
        .Value[3]   // P002 Manual setpoint
        .Value[4]   // P002 Flow setpoint
        .Value[5]   // P002 Linear Velocity setpoint
        .Value[6]   // Mixing Percentage setpoint
        .Value[7]   // Mixing Conductivity setpoint
   Membrane_Data : Membrane_Data := (Area := 19.38, Density := 1.01, NWP_TCF := 2.011, NWP_TCF_Temp := 22, NWP_TCF_Lookup_25[0] := 2.011, NWP_TCF_Lookup_25[1] := 1.943, NWP_TCF_Lookup_25[2] := 1.879, NWP_TCF_Lookup_25[3] := 1.818, NWP_TCF_Lookup_25[4] := 1.761, NWP_TCF_Lookup_25[5] := 1.706, NWP_TCF_Lookup_25[6] := 1.653, NWP_TCF_Lookup_25[7] := 1.604, NWP_TCF_Lookup_25[8] := 1.556, NWP_TCF_Lookup_25[9] := 1.511, NWP_TCF_Lookup_25[10] := 1.468, NWP_TCF_Lookup_25[11] := 1.426, NWP_TCF_Lookup_25[12] := 1.387, NWP_TCF_Lookup_25[13] := 1.349, NWP_TCF_Lookup_25[14] := 1.313, NWP_TCF_Lookup_25[15] := 1.278, NWP_TCF_Lookup_25[16] := 1.245, NWP_TCF_Lookup_25[17] := 1.213, NWP_TCF_Lookup_25[18] := 1.183, NWP_TCF_Lookup_25[19] := 1.154, NWP_TCF_Lookup_25[20] := 1.126, NWP_TCF_Lookup_25[21] := 1.099, NWP_TCF_Lookup_25[22] := 1.072, NWP_TCF_Lookup_25[23] := 1.047, NWP_TCF_Lookup_25[24] := 1.022, NWP_TCF_Lookup_25[25] := 1.0, NWP_TCF_Lookup_25[26] := 0.978, NWP_TCF_Lookup_25[27] := 0.956, NWP_TCF_Lookup_25[28] := 0.935, NWP_TCF_Lookup_25[29] := 0.915, NWP_TCF_Lookup_25[30] := 0.896, NWP_TCF_Lookup_25[31] := 0.877, NWP_TCF_Lookup_25[32] := 0.859, NWP_TCF_Lookup_25[33] := 0.841, NWP_TCF_Lookup_25[34] := 0.824, NWP_TCF_Lookup_25[35] := 0.808, NWP_TCF_Lookup_25[36] := 0.791, NWP_TCF_Lookup_25[37] := 0.777, NWP_TCF_Lookup_25[38] := 0.761, NWP_TCF_Lookup_25[39] := 0.747, NWP_TCF_Lookup_25[40] := 0.733, NWP_TCF_Lookup_25[41] := 0.719, NWP_TCF_Lookup_25[42] := 0.706, NWP_TCF_Lookup_25[43] := 0.694, NWP_TCF_Lookup_25[44] := 0.681, NWP_TCF_Lookup_25[45] := 0.669, NWP_TCF_Lookup_25[46] := 0.658, NWP_TCF_Lookup_25[47] := 0.646, NWP_TCF_Lookup_25[48] := 0.635, NWP_TCF_Lookup_25[49] := 0.624, NWP_TCF_Lookup_25[50] := 0.614, NWP_TCF_Lookup_25[51] := 0.604, NWP_TCF_Lookup_25[52] := 0.594);   // Membrane Data
   Memory_Data : Memory_Data := (Free_Mem_IO := 1022680, Free_Mem_DT := 276456, Free_Memory := 1299136, Total_Mem_IO := 1048576, Total_Mem_DT := 2097152, Total_Memory := 3145728, Biggest_IO_Mem_Size_Ava := 1021560, Biggest_DT_Mem_Size_Ava := 274976, Total_Mem_DT_Real := 2097152.0, Free_Mem_DT_Real := 276456.0, Used_Mem_DT_Real := 1820696.0, Percentage_Used_DT := 86.81755);
